(* IEC 61131-3 sources: volt/packages/volt-lsp-iec/test-corpus/lenze-mid/Device/Plc Logic/Application/Library Manager/L_OEEA_Library, 3.26.4.21 (Lenze), 47 files *)

(* ---- AXIS_REF_SIM.dut ---- *)
TYPE AXIS_REF_SIM :
STRUCT
	XENABLE : BOOL;
	XQUICKSTOP : BOOL;
	LRSETVELOCITY : LREAL;
	LRSETPOSITION : LREAL;
	XENABLED : BOOL;
	XREADY : BOOL;
	XDRIVEQSPACTIVE : BOOL;
	XERROR : BOOL;
	XWARNING : BOOL;
	EERRORID : L_IE1A_ErrorID;
	LRACTVELOCITY : LREAL;
	LRACTPOSITION : LREAL;
	XDIRECTIONPOSITIVE : BOOL;
	XDIRECTIONNEGATIVE : BOOL;
	DWDRIVEERRORID : DWORD;
	ETRAVERSINGRANGE : WORD := 1;
	LRCYCLELENGTH : LREAL := 560.0;
	LRFEEDCONSTANT : LREAL := 560.0;
	DWGEARNUMERATOR : DWORD := 77;
	DWGEARDENOMINATOR : DWORD := 6;
	XORIENTATION : BOOL := FALSE;
	EMCTRLMODE : DUT_eMctrlMode := 1;
	WNOOFHTLPERIODS : WORD := 128;
	DWHTLCOUNTERVALUE : DWORD;
	DWPOSRESOLUTION : DWORD := 65536;
	XTPRECEIVED : BOOL;
	LRTPLASTSCAN : LREAL;
	XSDOACTIVE : BOOL := TRUE;
	RDCBUSVOLTAGE : REAL;
	RMOTORCURRENT : REAL;
	RMOTORVOLTAGE : REAL;
	RMOTORSPEED : REAL;
	RMOTORFREQUENCY : REAL;
	DWERRORCODE : DWORD;
	RHEATSINKTEMP : REAL;
	RIXTLOAD : REAL;
	RIXT2LOAD : REAL;
	DWOPERATIONTIME : DWORD;
	DWSWITCHONTIME : DWORD;
	DWOPERATIONTIMECU : DWORD;
	DWOPERATIONTIMEFAN : DWORD;
END_STRUCT
END_TYPE

(* ---- DUT_EMCTRLMODE.dut ---- *)
TYPE DUT_EMCTRLMODE :
(
	OPENLOOP := 0,
	CLOSEDLOOP := 1
);
END_TYPE

(* ---- L_IE1A_ERRORID.dut ---- *)
TYPE L_IE1A_ERRORID :
(
	NOERROR := 0,
	MODULOAXISISREQUIRED := 17000,
	STARTPOSOUTOFCYCLELENGTH := 17003,
	CYCLELENGTHSHAVETOBEEQUAL := 17004,
	INVALIDDIRECTION := 17005,
	MARKSTACKLIMITREACHED := 17006,
	MAXMISSEDMARKS := 17007,
	INVALIDFOLLOWLINEACCVEL := 17008,
	INVALIDJOGGINGACCVEL := 17009,
	INVALIDSTOPDEC := 17010,
	INVALIDDIAMETER := 17011,
	TORQUEFOLLOWERNOTREADYFORMOTION := 17012,
	SPEEDFOLLOWERNOTREADYFORMOTION := 17013,
	INVALIDINVERTER := 17014,
	SDO_ACCESSFAILEDTOMOTORPARAMETERS := 17015,
	MISSEDMAPPINGPARAMETERLOWERSPEEDLIMIT := 17016,
	MISSEDMAPPINGPARAMETERUPPERSPEEDLIMIT := 17017,
	MISSEDMAPPINGPARAMETERTORQUEOFFSET := 17018,
	DANCERPOSOUTOFRANGE := 17019,
	INVALIDLIMITDANCERPOS := 17020,
	INVALIDCLUTCHPARAMETERS := 17021,
	WASNOTCALLEDDURINGMOTION := 17022,
	INVALIDNUMBEROFCAMPOINTS := 17030,
	INVALIDPATHPAR := 17032,
	INVALIDBLENDINGRADIUS := 17033,
	PATHNOTSUPPORTED := 17034,
	X_PATHLIMITPOSITIVEEXCEEDED := 17035,
	X_PATHLIMITNEGATIVEEXCEEDED := 17036,
	Y_PATHLIMITPOSITIVEEXCEEDED := 17037,
	Y_PATHLIMITNEGATIVEEXCEEDED := 17038,
	Z_PATHLIMITPOSITIVEEXCEEDED := 17039,
	Z_PATHLIMITNEGATIVEEXCEEDED := 17040,
	C_PATHLIMITPOSITIVEEXCEEDED := 17041,
	C_PATHLIMITNEGATIVEEXCEEDED := 17042,
	INVALIDPATHDATA := 17043,
	INVALIDTARGETPLC := 17047,
	MASTERISMOVING := 17100,
	INVALIDPODUCTLENGTH := 17101,
	TPSENSORNOTTEACHED := 17102,
	SLAVERECEIVEDGAPS := 17103,
	MASTERRECEIVEDGAPS := 17104,
	INTERNALERROR := 17105,
	INVALIDPARAMETERCUTTINGANGLE := 17106,
	INVALIDCUTTINGPARAMETERS := 17107,
	INVALIDCUTTINGLENGTH := 17108,
	SLAVENOTINPARKPOS := 17109,
	MASTERISREVERSING := 17110,
	INTINVALIDSELECTCAM := 17111,
	SELECTEDAXISISNOTSUPPORTED := 17112,
	AXISISNOTSUPPORTED := 17113,
	INVALIDPROFILE := 17114,
	AXISENABLEDISREQUIRED := 17115,
	CORRLIMITOUTOFCYCLELENGTH := 17116,
	CORRECTIONGREATERCORRWINDOW := 17117,
	INVALIDCNCPROGRAM := 17118,
	INVALIDGCODELINE := 17121,
	COORDSYSTEMACSNOTSUPPORTED := 17122,
	DANCERLIMITSNOTTEACHED := 17123,
	NOTREADYFORADDPROFILE := 17124,
	SLAVEPOSUPPERLIMIT := 17125,
	SLAVEPOSLOWERLIMIT := 17126,
	TARGETPOSUPPERLIMIT := 17127,
	INVALIDMARKPOSITION := 17128,
	INVALIDPOSITIONINGMODE := 17129,
	TEMPSENSORFAILURE := 17130,
	MAXCRITICALTEMPREACHED := 17131,
	INVALIDTEMPCONTROLPARAM := 17132,
	IDENTIFICATIONFAILED := 17133,
	PWMTASKCYCLEMISMATCH := 17134,
	CONCURRENTREQUESTTEMPCONTROL := 17135,
	TMNOTCALLEDINCYCLICTASK := 17136,
	TMDATABUSDISCONNECTED := 17137,
	INVALIDTMDATABUS := 17138,
	TMDATABUSCONFIGCHANGED := 17139,
	TMNOTCALLEDINMOTIONTASK := 17140,
	SLAVETMSTATESERVICE := 17141,
	COLLISIONDETECTIONDISABLED := 17142,
	COLLISIONDETECTED := 17143,
	INVALIDTMDATABUSORDER := 17144,
	CHANGEOFCONVEYORAXESNOTALLOWED := 17145,
	INVALIDSETTARGET := 17146,
	LOWERLIMITEXCEEDSUPPERLIMIT := 17147,
	SETTARGETSTACKLIMITREACHED := 17148,
	WORKPIECESTACKLIMITREACHED := 17149,
	INVALIDTRAVERSINGPROFILEPARAMETER := 17150,
	INVALIDTRAVERSINGCOILPARAMETER := 17151,
	TRAVERSINGANGULARSHIFTLIMITREACHED := 17152,
	AXESGROUPALREADYINUSE := 17153,
	UNDERVOLTAGEDCLINK := 17154,
	COUPLINGMODEREQUIRESMODULOAXIS := 17155,
	DUPLICATEDTM_ADDRESS := 17156,
	XAXISTMERROR := 17157,
	YAXISTMERROR := 17158,
	APAXISTMERROR := 17159,
	SLAVEXAXISTMERROR := 17160,
	SLAVEYAXISTMERROR := 17161,
	INVALIDMOVEPPACTIVE := 17162,
	INVALIDCONVEYORBELTPAR := 17163,
	IDENTIFICATIONDIAMETERFAILED := 17164,
	ACTDANCERPOSGTMAXDANCERPOS := 17165,
	INVALIDIDENTMAXDANCERPOS := 17166,
	INVALIDDANCERMATERIALLENGTH := 17167,
	LOADDIAMETERNOTALLOWED := 17168,
	INVALIDMASTERAXISREF := 17169,
	SYNCMODEVELACCREQUIRED := 17170,
	TEMPMAXCRITICALEXCEEDED := 17171,
	INVALIDTEMPCTRLPARAM := 17172,
	INVALIDSYNCSLAVEDIRECTION := 17173,
	MARKCORRECTIONINNEXTCYCLE := 17174,
	BASEVELOCITYNOTSUPPORTED := 17175,
	MOVEMENTBLOCKEDBYTRAINAHEAD := 17176,
	MARKDISTANCEGTZEROREQUIRED := 17177,
	INVALIDVIRTMASTERSETVELZERO := 17178,
	CONCURRENTMOTIONCMDDURINGHOMING := 17180,
	MISSINGMM_ADDRESS := 17901,
	TOOMANYMODULES := 17902,
	DUPLICATEDROOTMODULE := 17903,
	SLAVENOTFOUND := 17904,
	MISSINGAPPLICATIONREFERENCE := 17905,
	MISSINGMODULEREFERENCE := 17906,
	ERRORLISTOVERFLOW := 17907,
	ACDOWNSTRUCTINVALID := 17908,
	ACDSLAVESTRUCTINVALID := 17909,
	ACDSIZEOVERFLOW := 17910,
	COMPIDOUTOFRANGE := 17911,
	TOOMANYLEVELS := 17912,
	MMDSTRUCTINVALID := 17913,
	MODENUMBEROUTSIDERANGE := 18001,
	MODENUMBERNOTUSEDINCONFIG := 18002,
	MODECHANGENOTALLOWEDINCURRENTMODE := 18003,
	MODECHANGENOTALLOWEDINNEXTMODE := 18004,
	LI_MODENUMBEROUTSIDERANGE := 18005,
	LI_MODENUMBERNOTUSEDINCONFIG := 18006,
	LI_MODECHANGENOTALLOWEDREMOTE := 18007,
	LI_MODECHANGENOTALLOWEDINCURRENTMODE := 18008,
	LI_MODECHANGENOTALLOWEDINNEXTMODE := 18009,
	MORETHANONECOMMANDACTIVE := 18010,
	CONCURRENTCOMMAND := 18011,
	COMMANDNOTALLOWEDINCURRENTSTATE := 18012,
	LI_COMMANDSONLYINMODEPRODUCTION := 18013,
	LI_COMMANDNOTALLOWEDINREMOTE := 18014,
	LI_COMMANDNOTALLOWEDINCURRENTSTATE := 18015,
	DELAYTIMEINVALID_PT1FILTER := 19000,
	MODEINVALID_CURVE := 19002,
	MODEINVALID_COMPARE := 19003,
	MODEINVALID_CONVAXISV := 19005,
	DELAYTIMEINVALID_PROCESSCONTROLLER := 19006,
	RATETIMEINVALID_PROCESSCONTROLLER := 19007,
	RESETTIMEINVALID_PROCESSCONTROLLER := 19008,
	MODEINVALID_DELAY := 19024,
	ABORTEDBYSTARTIDENT_FRICTCOMP := 19030,
	ABORTEDBYFOLLOWERDISABLED_FRICTCOMP := 19031,
	MAXSPEEDNOTREACHED_FRICTCOMP := 19032,
	ACCTOOBIG_FRICTCOMP := 19033,
	DMINBIGGERDMAX_CALCDIAMETER := 19034,
	MAXSPEEDORMAXTORQUE_IDENTMINERTIA := 19048,
	ABORTEDBYSTARTIDENT_IDENTMINERTIA := 19049,
	ABORTEDBYFOLLOWERDISABLED_IDENTMINERTIA := 19050,
	ABORTEDBYFOLLOWERENABLED_IDENTMINERTIA := 19051,
	NMAXNOTREACHED_IDENTMINERTIA := 19052,
	MNOTREACHED_IDENTMINERTIA := 19053,
	MAXNROFTPEXCEEDED_MARKREGISTER := 19503,
	IDENTMODENOTSUPPORTED := 19801,
	MOTORRATEDSPEEDZERO := 19803,
	INERTIAMOTORZERO := 19804,
	STARTMODEINVALID := 19806,
	INVALIDEIGENFREQUENCY := 19807,
	INVALIDAMPLITUDERATIO := 19808,
	INVALIDOSCCOMPMODE := 19809,
	CHANGEOFOSCCOMPMODELOCKED := 19810,
	SDO_OTHERERROR := 20001,
	SDO_INVALIDINDEX := 20002,
	SDO_INVALIDOFFSET := 20003,
	SDO_INVALIDSIZE := 20004,
	SDO_INVALIDDATA := 20005,
	SDO_NOTREADY := 20006,
	SDO_BUSY := 20007,
	SDO_NOMEMORY := 20008,
	SDO_INVALIDPARM := 20009,
	SDO_INVALIDSTATE := 20010,
	SDO_TIMEOUT := 20011,
	SDO_INVALID_SLAVE_STATE := 20012,
	SDO_LINK_DISCONNECTED := 20013,
	SDO_ALL_CANNELS_BUSY := 20015,
	SDO_ABORTCODE_TOGGLE := 20020,
	SDO_ABORTCODE_TIMEOUT := 20021,
	SDO_ABORTCODE_CCS_SCS := 20022,
	SDO_ABORTCODE_BLK_SIZE := 20023,
	SDO_ABORTCODE_SEQNO := 20024,
	SDO_ABORTCODE_CRC := 20025,
	SDO_ABORTCODE_MEMORY := 20026,
	SDO_ABORTCODE_ACCESS := 20027,
	SDO_ABORTCODE_WRITEONLY := 20028,
	SDO_ABORTCODE_READONLY := 20029,
	SDO_ABORTCODE_INDEX := 20030,
	SDO_ABORTCODE_PDO_MAP := 20031,
	SDO_ABORTCODE_PDO_LEN := 20032,
	SDO_ABORTCODE_P_INCOMP := 20033,
	SDO_ABORTCODE_I_INCOMP := 20034,
	SDO_ABORTCODE_HARDWARE := 20035,
	SDO_ABORTCODE_DATA_SIZE := 20036,
	SDO_ABORTCODE_DATA_SIZE1 := 20037,
	SDO_ABORTCODE_DATA_SIZE2 := 20038,
	SDO_ABORTCODE_OFFSET := 20039,
	SDO_ABORTCODE_DATA_RANGE := 20040,
	SDO_ABORTCODE_DATA_RANGE1 := 20041,
	SDO_ABORTCODE_DATA_RANGE2 := 20042,
	SDO_ABORTCODE_MINMAX := 20043,
	SDO_ABORTCODE_GENERAL := 20044,
	SDO_ABORTCODE_TRANSFER := 20045,
	SDO_ABORTCODE_TRANSFER1 := 20046,
	SDO_ABORTCODE_TRANSFER2 := 20047,
	SDO_ABORTCODE_DICTIONARY := 20048,
	SDO_ABORTCODE_UNKNOWN := 20049,
	NOAXISREF := 20301,
	NOPARAMETER := 20302,
	NOVALIDPARAM := 20303,
	NOVALIDAXISSTATE := 20304,
	NOBOOLPARAM := 20305,
	SWLIMITPOS := 20306,
	SWLIMITNEG := 20307,
	NOVALID_MC_SOURCE := 20308,
	NOSETVALUESAVAILABLE := 20309,
	POWERFAILDURINGOPERATION := 20310,
	NOTREADYFORMOTION := 20311,
	POSSWLIMITREACHED := 20312,
	NEGSWLIMITREACHED := 20313,
	NOVALIDTPSOURCE := 20314,
	NOVALIDTPNUMBER := 20315,
	TPALREADYACTIVE := 20316,
	NOTTPSUPPORTED := 20317,
	NOTPACTIVE := 20318,
	NOEXTPINPUT := 20319,
	NOVALIDACCELERATION := 20320,
	NOVALIDDECELERATION := 20321,
	NOVALIDVELOCITY := 20322,
	ARITHMETICERROR := 20323,
	NOTAPPLICABLE := 20324,
	VELOCITYLIMITED := 20325,
	ACCELERATIONLIMITED := 20326,
	JERKLIMITED := 20327,
	TARGETOUTSIDESWLIMIT := 20328,
	NOVALIDACCELERATION_MOVEABSOLUTE := 20330,
	NOVALIDDECELERATION_MOVEABSOLUTE := 20331,
	NOVALIDVELOCITY_MOVEABSOLUTE := 20332,
	ARITHMETICERROR_MOVEABSOLUTE := 20333,
	NOTAPPLICABLE_MOVEABSOLUTE := 20334,
	VELOCITYLIMITED_MOVEABSOLUTE := 20335,
	ACCELERATIONLIMITED_MOVEABSOLUTE := 20336,
	JERKLIMITED_MOVEABSOLUTE := 20337,
	TARGETOUTSIDESWLIMIT_MOVEABSOLUTE := 20338,
	NOVALIDACCELERATION_MOVEADDITIVE := 20340,
	NOVALIDDECELERATION_MOVEADDITIVE := 20341,
	NOVALIDVELOCITY_MOVEADDITIVE := 20342,
	ARITHMETICERROR_MOVEADDITIVE := 20343,
	NOTAPPLICABLE_MOVEADDITIVE := 20344,
	VELOCITYLIMITED_MOVEADDITIVE := 20345,
	ACCELERATIONLIMITED_MOVEADDITIVE := 20346,
	JERKLIMITED_MOVEADDITIVE := 20347,
	TARGETOUTSIDESWLIMIT_MOVEADDITIVE := 20348,
	NOVALIDACCELERATION_MOVECONTAB := 20350,
	NOVALIDDECELERATION_MOVECONTAB := 20351,
	NOVALIDVELOCITY_MOVECONTAB := 20352,
	ARITHMETICERROR_MOVECONTAB := 20353,
	NOTAPPLICABLE_MOVECONTAB := 20354,
	VELOCITYLIMITED_MOVECONTAB := 20355,
	ACCELERATIONLIMITED_MOVECONTAB := 20356,
	JERKLIMITED_MOVECONTAB := 20357,
	TARGETOUTSIDESWLIMIT_MOVECONTAB := 20358,
	NOVALIDACCELERATION_MOVECONTREL := 20360,
	NOVALIDDECELERATION_MOVECONTREL := 20361,
	NOVALIDVELOCITY_MOVECONTREL := 20362,
	ARITHMETICERROR_MOVECONTREL := 20363,
	NOTAPPLICABLE_MOVECONTREL := 20364,
	VELOCITYLIMITED_MOVECONTREL := 20365,
	ACCELERATIONLIMITED_MOVECONTREL := 20366,
	JERKLIMITED_MOVECONTREL := 20367,
	TARGETOUTSIDESWLIMIT_MOVECONTREL := 20368,
	NOVALIDACCELERATION_MOVERELATIVE := 20370,
	NOVALIDDECELERATION_MOVERELATIVE := 20371,
	NOVALIDVELOCITY_MOVERELATIVE := 20372,
	ARITHMETICERROR_MOVERELATIVE := 20373,
	NOTAPPLICABLE_MOVERELATIVE := 20374,
	VELOCITYLIMITED_MOVERELATIVE := 20375,
	ACCELERATIONLIMITED_MOVERELATIVE := 20376,
	JERKLIMITED_MOVERELATIVE := 20377,
	TARGETOUTSIDESWLIMIT_MOVERELATIVE := 20378,
	NOVALIDACCELERATION_MOVESUPERIMP := 20380,
	NOVALIDDECELERATION_MOVESUPERIMP := 20381,
	NOVALIDVELOCITY_MOVESUPERIMP := 20382,
	ARITHMETICERROR_MOVESUPERIMP := 20383,
	NOTAPPLICABLE_MOVESUPERIMP := 20384,
	VELOCITYLIMITED_MOVESUPERIMP := 20385,
	ACCELERATIONLIMITED_MOVESUPERIMP := 20386,
	JERKLIMITED_MOVESUPERIMP := 20387,
	TARGETOUTSIDESWLIMIT_MOVESUPERIMP := 20388,
	NOVALIDACCELERATION_MOVEVELOCITY := 20390,
	NOVALIDDECELERATION_MOVEVELOCITY := 20391,
	NOVALIDVELOCITY_MOVEVELOCITY := 20392,
	ARITHMETICERROR_MOVEVELOCITY := 20393,
	NOTAPPLICABLE_MOVEVELOCITY := 20394,
	VELOCITYLIMITED_MOVEVELOCITY := 20395,
	ACCELERATIONLIMITED_MOVEVELOCITY := 20396,
	JERKLIMITED_MOVEVELOCITY := 20397,
	TARGETOUTSIDESWLIMIT_MOVEVELOCITY := 20398,
	NOVALIDDECELERATION_HALT := 20401,
	ARITHMETICERROR_HALT := 20403,
	ACCELERATIONLIMITED_HALT := 20406,
	JERKLIMITED_HALT := 20407,
	NOVALIDDECELERATION_STOP := 20411,
	ARITHMETICERROR_STOP := 20413,
	ACCELERATIONLIMITED_STOP := 20416,
	JERKLIMITED_STOP := 20417,
	NOVALIDDIRECTION := 20430,
	NOVALIDBUFFERMODE := 20431,
	DIRECTIONDISABLED := 20432,
	BLOCKEDBYAXISSTATE := 20433,
	NOVALIDOVERRIDE := 20434,
	CONCURRENT_MC_POWER := 20435,
	CONCURRENT_SETQUICKSTOP := 20436,
	DRIVE_PDO_INTERFACE_DISABLED := 20499,
	HWLIMITPOS := 20500,
	HWLIMITNEG := 20501,
	FOLLOWINGERROR1 := 20502,
	FOLLOWINGERROR2 := 20503,
	COMMUNICATIONFAIL := 20504,
	AXISINITFAIL := 20505,
	COMMTIMOUT := 20506,
	MASTERRESTARTFAIL := 20507,
	NOTREADYFORREINIT := 20508,
	ERRORDURINGINIT := 20509,
	SWITCHONNOTPOSSIBLE := 20510,
	DRIVEERROR := 20511,
	HOME_NOAUXPARAMETERS := 20512,
	HOME_MODENOTSUPPORTEDBYAXIS := 20513,
	HOME_MODEUNKNOWN := 20514,
	HOME_NOAUXTRIGGERINPUT := 20515,
	HOME_UNKNOWNTPCONFIG := 20516,
	HOME_WRITEHOMEPARAMETER := 20518,
	HOME_ERRORWHILEHOMING := 20519,
	HOME_ARITHMETICERROR := 20520,
	HOME_TORQUELIMNOTMAPPED := 20521,
	HOME_INVALIDVELACC := 20522,
	HOMETPEDGESETTINGNOTSUPPORTED := 20523,
	RESETDRIVEERRORFAILED := 20525,
	APPLICATIONERROR := 20526,
	APPLICATIONWARNING := 20527,
	BRAKE_POSITIONDRIFT := 20529,
	BRAKE_INVALIDMODE := 20530,
	BRAKE_TIMEOUTPRECONTROL := 20531,
	BRAKE_INVALIDBRAKESTATE := 20532,
	FAST_IO_OUT_WRONGOUTPUTSEL := 20533,
	FAST_IO_OUT_NOFREEENCODERAXIS := 20534,
	FAST_IO_OUT_FREEENCODERAXISWRONGPARAMETER := 20535,
	FAST_IO_OUT_MAPPINGFAULT := 20536,
	FAST_IO_OUT_FIFOOVERFLOW := 20537,
	TP_SELECT := 20538,
	TP_MODE := 20539,
	TP_EDGENOTAVAILABLE := 20541,
	TP_CHANNELNOTFREE := 20542,
	TP_MAPPINGFAULT := 20543,
	TP_INTERNALCHANNELNOTFREE := 20544,
	TP_TIMEOUT := 20545,
	TP_COMMUNICATIONERROR := 20546,
	TP_SIGNAL := 20547,
	TP_NOFREEENCODERAXIS := 20548,
	TP_PARAMETERRISINGEDGEWRONGVALUE := 20550,
	TP_PARAMETERFALLINGRISINGEDGEWRONGVALUE := 20551,
	TP_INTERNALERROR := 20552,
	SETVALUESGTMAXAPPVALUES := 20600,
	SETVALUESINCONSISTENT := 20601,
	POSDIFFGTHALFCYCLELENGTH := 20602,
	INVALIDTASKCYCLETIME := 20603,
	INIT_WRITEERRORSDO := 20650,
	INIT_READERRORSDO := 20651,
	INIT_MAXTASKTIME := 20652,
	INIT_TORQUEREFISZERO := 20653,
	INIT_MOTORRATEDSPEEDISZERO := 20654,
	INIT_REVISIONNOTVALID := 20655,
	INIT_ENCCOUNTNOTVALID := 20656,
	INIT_ENCREVNOTVALID := 20657,
	INIT_ENCCRCNOTVALID := 20658,
	INIT_ENCABSPOSNOTAVAILABLE := 20659,
	CONTROLLERFIRMWARENOTCOMPATIBLE := 20660,
	INVALIDMODE := 20661,
	ENCBPB_INIT_FAILED := 20662,
	LEDNOTSUPPORTEDBYDEVICE := 20663,
	INVALIDGEARFACTOR := 20664,
	POSOUTOFCYCLELENGTH := 20665,
	CYCLELENGTHINVALID_ADDOFFSETCYCLIC := 20666,
	POSININVALID_ADDOFFSETCYCLIC := 20667,
	CYCLELENGTHINVALID_ZERODETECT := 20668,
	POSININVALID_ZERODETECT := 20669,
	STARTPOSINVALID_INTEGRATEAXIS := 20670,
	INVALIDINPUTJOGPOSJOGNEG := 20671,
	VALUEOUTOFRANGE := 20672,
	STATENOTEQUALDISABLED := 20673,
	INVALIDINPUT_BRAKETEST := 20674,
	ALREADYACTIVE_BRAKETEST := 20675,
	INVALIDINPUT_BRAKEGRINDIN := 20676,
	ALREADYACTIVE_GRINDIN := 20677,
	INVALIDCONTROLMODE := 20678,
	VIRTUALAXISNOTSUPPORTED := 20679,
	AXISNOTDISABLED := 20680,
	INVALIDFEEDCONSTANT := 20681,
	INVALIDTRAVERSINGRANGE := 20682,
	INVALIDCYCLELENGTH := 20683,
	INVALIDPOSRESOLUTION := 20684,
	TORQUELIMTOOLARGE := 20685,
	TORQUELIMLESSTHANZERO := 20686,
	ENCSIGNALINVALID := 20687,
	ENCSIGNALGTMEASURINGRANGE := 20688,
	INVALIDENCMEASURINGRANGE := 20689,
	DRIVESTOACTIVE := 20690,
	DRIVECINHACTIVE := 20691,
	INVALIDSWLIMITS := 20692,
	NOVALIDJERK := 20693,
	MISSEDMAPPINGPARAMETERVLTARGETVEL := 20694,
	MISSEDMAPPINGPARAMETERVLACTUALVEL := 20695,
	AXISNOTHOMED := 20696,
	AXISNOTINSIMPLEMODE := 20697,
	AXISINSIMPLEMODE := 20698,
	FUNCTIONNOTSUPPORTEDBYAXIS := 20699,
	EXECUTIONINDEXALREADYINUSE := 20700,
	SS1ACTIVE := 20701,
	SS2ACTIVE := 20702,
	VELOCITYLIMITEDBYSLS1 := 20703,
	VELOCITYLIMITEDBYSLS2 := 20704,
	VELOCITYLIMITEDBYSLS3 := 20705,
	VELOCITYLIMITEDBYSLS4 := 20706,
	INVALIDEXECUTIONINDEX := 20707,
	INVALIDFILTERDEPTH := 20708,
	PARAMSETFAILEDJOGVEL := 20709,
	PARAMSETFAILEDJOGACC := 20710,
	PARAMSETFAILEDJOGDEC := 20711,
	PARAMSETFAILEDJOGJERK := 20712,
	PARAMSETFAILEDHALTDEC := 20713,
	PARAMSETFAILEDHALTJERK := 20714,
	PARAMSETFAILEDQSPAPPLDEC := 20715,
	PARAMSETFAILEDQSPAPPLJERK := 20716,
	PARAMSETFAILEDHOMEPOSITION := 20717,
	PARAMSETFAILEDHOMEMODE := 20718,
	PARAMSETFAILEDHOMESTOPMODE := 20719,
	PARAMSETFAILEDHOMETARGETPOSITION := 20720,
	PARAMSETFAILEDHOMEVELOCITY1 := 20721,
	PARAMSETFAILEDHOMEVELOCITY2 := 20722,
	PARAMSETFAILEDHOMEACCELERATION1 := 20723,
	PARAMSETFAILEDHOMEACCELERATION2 := 20724,
	PARAMSETFAILEDHOMEJERK := 20725,
	PARAMSETFAILEDHOMETORQUELIMIT := 20726,
	PARAMSETFAILEDHOMETORQUETIME := 20727,
	PARAMSETFAILEDHOMETPCONFIG := 20728,
	PARAMSETFAILEDDRIVEHOMEMODE := 20729,
	PARAMREADFAILED := 20730,
	PARAMROLLBACKFAILED := 20731,
	POSCTRLNOTSUPPORTED := 20732,
	TORQUECTRLNOTSUPPORTED := 20733,
	SETPOSITIONINPDOREQUIRED := 20734,
	SETVELOCITYINPDOREQUIRED := 20735,
	SETTORQUEINPDOREQUIRED := 20736,
	UPPERSPEEDLIMINPDOREQUIRED := 20737,
	LOWERSPEEDLIMINPDOREQUIRED := 20738,
	ACTPOSITIONINPDOREQUIRED := 20739,
	BRAKEGRINDININVALIDPOSITIONLIMITS := 20740,
	BRAKEGRINDINSTARTPOSOUTSIDEPOSLIM := 20741,
	BRAKEGRINDINDISTANCENOTSUFFICIENT := 20742,
	SAFETYNOTSUPPORTEDBYDRIVE := 20743,
	SAFETYCONTROLWORDINPDOREQUIRED := 20744,
	SETPOSITIONONSLAVEAXISNOTALLOWED := 20745,
	ENCODERVELOCITYGTMAXVELOCITY := 20746,
	INVALIDENCODERSIGNAL := 20747,
	DRIVESAFEBRAKECTRLACTIVE := 20748,
	POSRECONSTRDATAINKONSISTENT := 20750,
	POSRECONSTRHOMEPOSAVAILABLENOTACTIVE := 20751,
	POSRECONSTRNOTACTIVATED := 20752,
	POSRECONSTRAXISWASVIRTUAL := 20753,
	POSRECONSTRORIENTATIONCHANGED := 20754,
	POSRECONSTRTRAVERSINGRANGECHANGED := 20755,
	POSRECONSTRCYCLELENGTHCHANGED := 20756,
	POSRECONSTRUNITFACTORCHANGED := 20757,
	POSRECONSTRRESETBYENCERROR := 20758,
	POSRECONSTRRESETBYFDBCHANGED := 20759,
	POSRECONSTRENCCRCCHANGED := 20760,
	POSRECONSTRNOFDBPOSAVAILABLE := 20761,
	POSRECONSTRABSENCREQUIRED := 20762,
	POSRECONSTRDATAVERSIONCHANGED := 20763,
	POSRECONSTRNODATAAVAILABLE := 20764,
	POSRECONSTRNOMEMORYAVAILABLE := 20765,
	POSRECONSTRPOSOUTSIDERESTORETRESHOLD := 20766,
	POSRECONSTRRESETBYFDBOPENCIRC := 20767,
	MAINAXISNOTREADY := 21001,
	GROUPSTATEUNDEFINED := 21002,
	AXISDISABLED := 21003,
	TRANSFORMATIONERROR := 21004,
	AXISINERRORSTOP := 21005,
	AXISLIMITVIOLATIONMAINAXIS := 21006,
	AXISLIMITVIOLATIONREALAXIS := 21007,
	AXISLIMITVIOLATIONPASSIVEAXIS := 21008,
	REALAXISDISABLED := 21009,
	NOVALIDPATHCOICE_MOVECIRCABS := 21010,
	NOVALIDCIRCMODE_MOVECIRCABS := 21011,
	NOVALIDTRANSITIONPARAMETER_MOVECIRCABS := 21012,
	NOVALIDVELOCITY_MOVECIRCABS := 21013,
	NOVALIDACCELERATION_MOVECIRCABS := 21014,
	NOVALIDDECELERATION_MOVECIRCABS := 21015,
	NOVALIDJERK_MOVECIRCABS := 21016,
	TARGETOUTSIDESWLIMITSPASSIVEJOINTS_MOVECIRCABS := 21017,
	TARGETOUTSIDESWLIMITSMAINAXISX_MOVECIRCABS := 21018,
	TARGETOUTSIDESWLIMITSMAINAXISY_MOVECIRCABS := 21019,
	TARGETOUTSIDESWLIMITSMAINAXISZ_MOVECIRCABS := 21020,
	TARGETOUTSIDESWLIMITSMAINAXISA_MOVECIRCABS := 21021,
	TARGETOUTSIDESWLIMITSMAINAXISB_MOVECIRCABS := 21022,
	TARGETOUTSIDESWLIMITSMAINAXISC_MOVECIRCABS := 21023,
	TARGETOUTSIDESWLIMITSREALAXIS1_MOVECIRCABS := 21024,
	TARGETOUTSIDESWLIMITSREALAXIS2_MOVECIRCABS := 21025,
	TARGETOUTSIDESWLIMITSREALAXIS3_MOVECIRCABS := 21026,
	TARGETOUTSIDESWLIMITSREALAXIS4_MOVECIRCABS := 21027,
	TARGETOUTSIDESWLIMITSREALAXIS5_MOVECIRCABS := 21028,
	TARGETOUTSIDESWLIMITSREALAXIS6_MOVECIRCABS := 21029,
	TARGETOUTSIDESWLIMITSAUXAXIS1_MOVECIRCABS := 21030,
	TARGETOUTSIDESWLIMITSAUXAXIS2_MOVECIRCABS := 21031,
	TARGETOUTSIDESWLIMITSAUXAXIS3_MOVECIRCABS := 21032,
	TARGETOUTSIDESWLIMITSAUXAXIS4_MOVECIRCABS := 21033,
	TARGETOUTSIDESWLIMITSAUXAXIS5_MOVECIRCABS := 21034,
	TARGETOUTSIDESWLIMITSAUXAXIS6_MOVECIRCABS := 21035,
	TARGETTRANSFORMATIONERROR_MOVECIRCABS := 21036,
	TARGETSINGULARPOS_MOVECIRCABS := 21037,
	BORDEROUTSIDESWLIMITSPASSIVEJOINTS_MOVECIRCABS := 21038,
	BORDEROUTSIDESWLIMITSMAINAXISX_MOVECIRCABS := 21039,
	BORDEROUTSIDESWLIMITSMAINAXISY_MOVECIRCABS := 21040,
	BORDEROUTSIDESWLIMITSMAINAXISZ_MOVECIRCABS := 21041,
	BORDEROUTSIDESWLIMITSMAINAXISA_MOVECIRCABS := 21042,
	BORDEROUTSIDESWLIMITSMAINAXISB_MOVECIRCABS := 21043,
	BORDEROUTSIDESWLIMITSMAINAXISC_MOVECIRCABS := 21044,
	BORDEROUTSIDESWLIMITSREALAXIS1_MOVECIRCABS := 21045,
	BORDEROUTSIDESWLIMITSREALAXIS2_MOVECIRCABS := 21046,
	BORDEROUTSIDESWLIMITSREALAXIS3_MOVECIRCABS := 21047,
	BORDEROUTSIDESWLIMITSREALAXIS4_MOVECIRCABS := 21048,
	BORDEROUTSIDESWLIMITSREALAXIS5_MOVECIRCABS := 21049,
	BORDEROUTSIDESWLIMITSREALAXIS6_MOVECIRCABS := 21050,
	BORDEROUTSIDESWLIMITSAUXAXIS1_MOVECIRCABS := 21051,
	BORDEROUTSIDESWLIMITSAUXAXIS2_MOVECIRCABS := 21052,
	BORDEROUTSIDESWLIMITSAUXAXIS3_MOVECIRCABS := 21053,
	BORDEROUTSIDESWLIMITSAUXAXIS4_MOVECIRCABS := 21054,
	BORDEROUTSIDESWLIMITSAUXAXIS5_MOVECIRCABS := 21055,
	BORDEROUTSIDESWLIMITSAUXAXIS6_MOVECIRCABS := 21056,
	BORDERTRANSFORMATIONERROR_MOVECIRCABS := 21057,
	BORDERSINGULARPOS_MOVECIRCABS := 21058,
	ILLEGALPARAMETER_MOVECIRCABS := 21059,
	NOVALIDPATHCOICE_MOVECIRCREL := 21060,
	NOVALIDCIRCMODE_MOVECIRCREL := 21061,
	NOVALIDTRANSITIONPARAMETER_MOVECIRCREL := 21062,
	NOVALIDVELOCITY_MOVECIRCREL := 21063,
	NOVALIDACCELERATION_MOVECIRCREL := 21064,
	NOVALIDDECELERATION_MOVECIRCREL := 21065,
	NOVALIDJERK_MOVECIRCREL := 21066,
	TARGETOUTSIDESWLIMITSPASSIVEJOINTS_MOVECIRCREL := 21067,
	TARGETOUTSIDESWLIMITSMAINAXISX_MOVECIRCREL := 21068,
	TARGETOUTSIDESWLIMITSMAINAXISY_MOVECIRCREL := 21069,
	TARGETOUTSIDESWLIMITSMAINAXISZ_MOVECIRCREL := 21070,
	TARGETOUTSIDESWLIMITSMAINAXISA_MOVECIRCREL := 21071,
	TARGETOUTSIDESWLIMITSMAINAXISB_MOVECIRCREL := 21072,
	TARGETOUTSIDESWLIMITSMAINAXISC_MOVECIRCREL := 21073,
	TARGETOUTSIDESWLIMITSREALAXIS1_MOVECIRCREL := 21074,
	TARGETOUTSIDESWLIMITSREALAXIS2_MOVECIRCREL := 21075,
	TARGETOUTSIDESWLIMITSREALAXIS3_MOVECIRCREL := 21076,
	TARGETOUTSIDESWLIMITSREALAXIS4_MOVECIRCREL := 21077,
	TARGETOUTSIDESWLIMITSREALAXIS5_MOVECIRCREL := 21078,
	TARGETOUTSIDESWLIMITSREALAXIS6_MOVECIRCREL := 21079,
	TARGETOUTSIDESWLIMITSAUXAXIS1_MOVECIRCREL := 21080,
	TARGETOUTSIDESWLIMITSAUXAXIS2_MOVECIRCREL := 21081,
	TARGETOUTSIDESWLIMITSAUXAXIS3_MOVECIRCREL := 21082,
	TARGETOUTSIDESWLIMITSAUXAXIS4_MOVECIRCREL := 21083,
	TARGETOUTSIDESWLIMITSAUXAXIS5_MOVECIRCREL := 21084,
	TARGETOUTSIDESWLIMITSAUXAXIS6_MOVECIRCREL := 21085,
	TARGETTRANSFORMATIONERROR_MOVECIRCREL := 21086,
	TARGETSINGULARPOS_MOVECIRCREL := 21087,
	BORDEROUTSIDESWLIMITSPASSIVEJOINTS_MOVECIRCREL := 21088,
	BORDEROUTSIDESWLIMITSMAINAXISX_MOVECIRCREL := 21089,
	BORDEROUTSIDESWLIMITSMAINAXISY_MOVECIRCREL := 21090,
	BORDEROUTSIDESWLIMITSMAINAXISZ_MOVECIRCREL := 21091,
	BORDEROUTSIDESWLIMITSMAINAXISA_MOVECIRCREL := 21092,
	BORDEROUTSIDESWLIMITSMAINAXISB_MOVECIRCREL := 21093,
	BORDEROUTSIDESWLIMITSMAINAXISC_MOVECIRCREL := 21094,
	BORDEROUTSIDESWLIMITSREALAXIS1_MOVECIRCREL := 21095,
	BORDEROUTSIDESWLIMITSREALAXIS2_MOVECIRCREL := 21096,
	BORDEROUTSIDESWLIMITSREALAXIS3_MOVECIRCREL := 21097,
	BORDEROUTSIDESWLIMITSREALAXIS4_MOVECIRCREL := 21098,
	BORDEROUTSIDESWLIMITSREALAXIS5_MOVECIRCREL := 21099,
	BORDEROUTSIDESWLIMITSREALAXIS6_MOVECIRCREL := 21100,
	BORDEROUTSIDESWLIMITSAUXAXIS1_MOVECIRCREL := 21101,
	BORDEROUTSIDESWLIMITSAUXAXIS2_MOVECIRCREL := 21102,
	BORDEROUTSIDESWLIMITSAUXAXIS3_MOVECIRCREL := 21103,
	BORDEROUTSIDESWLIMITSAUXAXIS4_MOVECIRCREL := 21104,
	BORDEROUTSIDESWLIMITSAUXAXIS5_MOVECIRCREL := 21105,
	BORDEROUTSIDESWLIMITSAUXAXIS6_MOVECIRCREL := 21106,
	BORDERTRANSFORMATIONERROR_MOVECIRCREL := 21107,
	BORDERSINGULARPOS_MOVECIRCREL := 21108,
	ILLEGALPARAMETER_MOVECIRCREL := 21109,
	NOVALIDTRANSITIONPARAMETER_MOVELINABS := 21110,
	NOVALIDVELOCITY_MOVELINABS := 21111,
	NOVALIDACCELERATION_MOVELINABS := 21112,
	NOVALIDDECELERATION_MOVELINABS := 21113,
	NOVALIDJERK_MOVELINABS := 21114,
	TARGETOUTSIDESWLIMITSPASSIVEJOINTS_MOVELINABS := 21115,
	TARGETOUTSIDESWLIMITSMAINAXISX_MOVELINABS := 21116,
	TARGETOUTSIDESWLIMITSMAINAXISY_MOVELINABS := 21117,
	TARGETOUTSIDESWLIMITSMAINAXISZ_MOVELINABS := 21118,
	TARGETOUTSIDESWLIMITSMAINAXISA_MOVELINABS := 21119,
	TARGETOUTSIDESWLIMITSMAINAXISB_MOVELINABS := 21120,
	TARGETOUTSIDESWLIMITSMAINAXISC_MOVELINABS := 21121,
	TARGETOUTSIDESWLIMITSREALAXIS1_MOVELINABS := 21122,
	TARGETOUTSIDESWLIMITSREALAXIS2_MOVELINABS := 21123,
	TARGETOUTSIDESWLIMITSREALAXIS3_MOVELINABS := 21124,
	TARGETOUTSIDESWLIMITSREALAXIS4_MOVELINABS := 21125,
	TARGETOUTSIDESWLIMITSREALAXIS5_MOVELINABS := 21126,
	TARGETOUTSIDESWLIMITSREALAXIS6_MOVELINABS := 21127,
	TARGETOUTSIDESWLIMITSAUXAXIS1_MOVELINABS := 21128,
	TARGETOUTSIDESWLIMITSAUXAXIS2_MOVELINABS := 21129,
	TARGETOUTSIDESWLIMITSAUXAXIS3_MOVELINABS := 21130,
	TARGETOUTSIDESWLIMITSAUXAXIS4_MOVELINABS := 21131,
	TARGETOUTSIDESWLIMITSAUXAXIS5_MOVELINABS := 21132,
	TARGETOUTSIDESWLIMITSAUXAXIS6_MOVELINABS := 21133,
	TARGETTRANSFORMATIONERROR_MOVELINABS := 21134,
	TARGETSINGULARPOS_MOVELINABS := 21135,
	ILLEGALPARAMETER_MOVELINABS := 21136,
	NOVALIDTRANSITIONPARAMETER_MOVELINREL := 21137,
	NOVALIDVELOCITY_MOVELINREL := 21138,
	NOVALIDACCELERATION_MOVELINREL := 21139,
	NOVALIDDECELERATION_MOVELINREL := 21140,
	NOVALIDJERK_MOVELINREL := 21141,
	TARGETOUTSIDESWLIMITSPASSIVEJOINTS_MOVELINREL := 21142,
	TARGETOUTSIDESWLIMITSMAINAXISX_MOVELINREL := 21143,
	TARGETOUTSIDESWLIMITSMAINAXISY_MOVELINREL := 21144,
	TARGETOUTSIDESWLIMITSMAINAXISZ_MOVELINREL := 21145,
	TARGETOUTSIDESWLIMITSMAINAXISA_MOVELINREL := 21146,
	TARGETOUTSIDESWLIMITSMAINAXISB_MOVELINREL := 21147,
	TARGETOUTSIDESWLIMITSMAINAXISC_MOVELINREL := 21148,
	TARGETOUTSIDESWLIMITSREALAXIS1_MOVELINREL := 21149,
	TARGETOUTSIDESWLIMITSREALAXIS2_MOVELINREL := 21150,
	TARGETOUTSIDESWLIMITSREALAXIS3_MOVELINREL := 21151,
	TARGETOUTSIDESWLIMITSREALAXIS4_MOVELINREL := 21152,
	TARGETOUTSIDESWLIMITSREALAXIS5_MOVELINREL := 21153,
	TARGETOUTSIDESWLIMITSREALAXIS6_MOVELINREL := 21154,
	TARGETOUTSIDESWLIMITSAUXAXIS1_MOVELINREL := 21155,
	TARGETOUTSIDESWLIMITSAUXAXIS2_MOVELINREL := 21156,
	TARGETOUTSIDESWLIMITSAUXAXIS3_MOVELINREL := 21157,
	TARGETOUTSIDESWLIMITSAUXAXIS4_MOVELINREL := 21158,
	TARGETOUTSIDESWLIMITSAUXAXIS5_MOVELINREL := 21159,
	TARGETOUTSIDESWLIMITSAUXAXIS6_MOVELINREL := 21160,
	TARGETTRANSFORMATIONERROR_MOVELINREL := 21161,
	TARGETSINGULARPOS_MOVELINREL := 21162,
	ILLEGALPARAMETER_MOVELINREL := 21163,
	NOVALIDTRANSITIONPARAMETER_MOVEDIRABS := 21164,
	NOVALIDVELOCITY_MOVEDIRABS := 21165,
	NOVALIDACCELERATION_MOVEDIRABS := 21166,
	NOVALIDDECELERATION_MOVEDIRABS := 21167,
	NOVALIDJERK_MOVEDIRABS := 21168,
	TARGETOUTSIDESWLIMITSPASSIVEJOINTS_MOVEDIRABS := 21169,
	TARGETOUTSIDESWLIMITSMAINAXISX_MOVEDIRABS := 21170,
	TARGETOUTSIDESWLIMITSMAINAXISY_MOVEDIRABS := 21171,
	TARGETOUTSIDESWLIMITSMAINAXISZ_MOVEDIRABS := 21172,
	TARGETOUTSIDESWLIMITSMAINAXISA_MOVEDIRABS := 21173,
	TARGETOUTSIDESWLIMITSMAINAXISB_MOVEDIRABS := 21174,
	TARGETOUTSIDESWLIMITSMAINAXISC_MOVEDIRABS := 21175,
	TARGETOUTSIDESWLIMITSREALAXIS1_MOVEDIRABS := 21176,
	TARGETOUTSIDESWLIMITSREALAXIS2_MOVEDIRABS := 21177,
	TARGETOUTSIDESWLIMITSREALAXIS3_MOVEDIRABS := 21178,
	TARGETOUTSIDESWLIMITSREALAXIS4_MOVEDIRABS := 21179,
	TARGETOUTSIDESWLIMITSREALAXIS5_MOVEDIRABS := 21180,
	TARGETOUTSIDESWLIMITSREALAXIS6_MOVEDIRABS := 21181,
	TARGETOUTSIDESWLIMITSAUXAXIS1_MOVEDIRABS := 21182,
	TARGETOUTSIDESWLIMITSAUXAXIS2_MOVEDIRABS := 21183,
	TARGETOUTSIDESWLIMITSAUXAXIS3_MOVEDIRABS := 21184,
	TARGETOUTSIDESWLIMITSAUXAXIS4_MOVEDIRABS := 21185,
	TARGETOUTSIDESWLIMITSAUXAXIS5_MOVEDIRABS := 21186,
	TARGETOUTSIDESWLIMITSAUXAXIS6_MOVEDIRABS := 21187,
	TARGETTRANSFORMATIONERROR_MOVEDIRABS := 21188,
	ILLEGALPARAMETER_MOVEDIRABS := 21189,
	NOVALIDTRANSITIONPARAMETER_MOVEDIRREL := 21190,
	NOVALIDVELOCITY_MOVEDIRREL := 21191,
	NOVALIDACCELERATION_MOVEDIRREL := 21192,
	NOVALIDDECELERATION_MOVEDIRREL := 21193,
	NOVALIDJERK_MOVEDIRREL := 21194,
	TARGETOUTSIDESWLIMITSPASSIVEJOINTS_MOVEDIRREL := 21195,
	TARGETOUTSIDESWLIMITSMAINAXISX_MOVEDIRREL := 21196,
	TARGETOUTSIDESWLIMITSMAINAXISY_MOVEDIRREL := 21197,
	TARGETOUTSIDESWLIMITSMAINAXISZ_MOVEDIRREL := 21198,
	TARGETOUTSIDESWLIMITSMAINAXISA_MOVEDIRREL := 21199,
	TARGETOUTSIDESWLIMITSMAINAXISB_MOVEDIRREL := 21200,
	TARGETOUTSIDESWLIMITSMAINAXISC_MOVEDIRREL := 21201,
	TARGETOUTSIDESWLIMITSREALAXIS1_MOVEDIRREL := 21202,
	TARGETOUTSIDESWLIMITSREALAXIS2_MOVEDIRREL := 21203,
	TARGETOUTSIDESWLIMITSREALAXIS3_MOVEDIRREL := 21204,
	TARGETOUTSIDESWLIMITSREALAXIS4_MOVEDIRREL := 21205,
	TARGETOUTSIDESWLIMITSREALAXIS5_MOVEDIRREL := 21206,
	TARGETOUTSIDESWLIMITSREALAXIS6_MOVEDIRREL := 21207,
	TARGETOUTSIDESWLIMITSAUXAXIS1_MOVEDIRREL := 21208,
	TARGETOUTSIDESWLIMITSAUXAXIS2_MOVEDIRREL := 21209,
	TARGETOUTSIDESWLIMITSAUXAXIS3_MOVEDIRREL := 21210,
	TARGETOUTSIDESWLIMITSAUXAXIS4_MOVEDIRREL := 21211,
	TARGETOUTSIDESWLIMITSAUXAXIS5_MOVEDIRREL := 21212,
	TARGETOUTSIDESWLIMITSAUXAXIS6_MOVEDIRREL := 21213,
	TARGETTRANSFORMATIONERROR_MOVEDIRREL := 21214,
	ILLEGALPARAMETER_MOVEDIRREL := 21215,
	NOVALIDVELOCITY_MANMODE := 21216,
	NOVALIDACCELERATION_MANMODE := 21217,
	NOVALIDDECELERATION_MANMODE := 21218,
	NOVALIDJERK_MANMODE := 21219,
	MANUALMODEILLEGALPARAMETER := 21220,
	KINEMATICILLEGALPARAMETER := 21221,
	AXESGROUPINERRORSTOP := 21222,
	TOOLINUSE := 21223,
	INVALIDTOOL := 21224,
	AXESGROUPINMOVEMENT := 21225,
	INVALIDCOORDSYSTEM := 21226,
	AXISEXTERNALENABLED := 21227,
	UNSUPPORTEDCOORDSYSTEM := 21228,
	REALAXISNOTREADY := 21229,
	INVALIDAXESGROUPSTATE := 21230,
	REALAXISOUTSIDEWORKINGRANGE := 21231,
	SINGULARPOSITION := 21232,
	L_MC4P_INTERNALERROR := 21233,
	AXESGROUPEXTERNALSTOPPING := 21234,
	RESETAXESGROUPERRORFAILED := 21237,
	ILLEGALTEACHPOSITION := 21238,
	NOTENOUGHMEMORYPATHDATALIST := 21239,
	NOVALIDROTATIONVELOCITY_MOVECIRCABS := 21240,
	NOVALIDROTATIONACCELERATION_MOVECIRCABS := 21241,
	NOVALIDROTATIONJERK_MOVECIRCABS := 21242,
	NOVALIDROTATIONVELOCITY_MOVECIRCREL := 21243,
	NOVALIDROTATIONACCELERATION_MOVECIRCREL := 21244,
	NOVALIDROTATIONJERK_MOVECIRCREL := 21245,
	NOVALIDROTATIONVELOCITY_MOVELINABS := 21246,
	NOVALIDROTATIONACCELERATION_MOVELINABS := 21247,
	NOVALIDROTATIONJERK_MOVELINABS := 21248,
	NOVALIDROTATIONVELOCITY_MOVELINREL := 21249,
	NOVALIDROTATIONACCELERATION_MOVELINREL := 21250,
	NOVALIDROTATIONJERK_MOVELINREL := 21251,
	PATHLIMITVIOLATION_MOVELINABS := 21252,
	PATHLIMITVIOLATION_MOVELINREL := 21253,
	PATHLIMITVIOLATION_MOVECIRCABS := 21254,
	PATHLIMITVIOLATION_MOVECIRCREL := 21255,
	PATHLIMITVIOLATION_MOVEDIRABS := 21256,
	PATHLIMITVIOLATION_MOVEDIRREL := 21257,
	AXISGROUPNOTHOMED := 21258,
	MAINAXISTYPEMODULONOTALLOWED := 21259,
	AXISTYPEMODULONOTALLOWED := 21260,
	AXISLIMITVIOLATIONREALAXIS1VELOCITY := 21261,
	AXISLIMITVIOLATIONREALAXIS2VELOCITY := 21262,
	AXISLIMITVIOLATIONREALAXIS3VELOCITY := 21263,
	AXISLIMITVIOLATIONREALAXIS4VELOCITY := 21264,
	AXISLIMITVIOLATIONREALAXIS5VELOCITY := 21265,
	AXISLIMITVIOLATIONREALAXIS6VELOCITY := 21266,
	AXISLIMITVIOLATIONREALAXIS1ACCELERATION := 21267,
	AXISLIMITVIOLATIONREALAXIS2ACCELERATION := 21268,
	AXISLIMITVIOLATIONREALAXIS3ACCELERATION := 21269,
	AXISLIMITVIOLATIONREALAXIS4ACCELERATION := 21270,
	AXISLIMITVIOLATIONREALAXIS5ACCELERATION := 21271,
	AXISLIMITVIOLATIONREALAXIS6ACCELERATION := 21272,
	AUXAXISSEQUENCEINVALID := 21273,
	AUXAXISNOTALLOWED := 21274,
	ILLEGALTRACKINGPARAMETER := 21275,
	SYNCHRONISATIONERROR := 21276,
	PCSINUSE := 21277,
	TRACKINGFBNOTCALLED := 21278,
	MASTERAXISNOTREADY := 21279,
	MOVEDIRECTNOTALLOWED := 21280,
	AUXAXISNOVALIDVELOCITY := 21281,
	AUXAXISNOVALIDACCELERATION := 21282,
	AUXAXISNOVALIDJERK := 21283,
	MAINAXISNOTCONNECTED := 21284,
	REALAXISNOTCONNECTED := 21285,
	AXESGROUPNOTINITIALIZED := 21286,
	DISABLEDBYPARAMETERTRANSFER := 21287,
	REALAXIS1_ALREADYINUSE := 21288,
	REALAXIS2_ALREADYINUSE := 21289,
	REALAXIS3_ALREADYINUSE := 21290,
	REALAXIS4_ALREADYINUSE := 21291,
	REALAXIS5_ALREADYINUSE := 21292,
	REALAXIS6_ALREADYINUSE := 21293,
	AUXAXIS1_ALREADYINUSE := 21294,
	AUXAXIS2_ALREADYINUSE := 21295,
	AUXAXIS3_ALREADYINUSE := 21296,
	AUXAXIS4_ALREADYINUSE := 21297,
	AUXAXIS5_ALREADYINUSE := 21298,
	AUXAXIS6_ALREADYINUSE := 21299,
	NOVALIDTRANSITIONMODE_MOVECIRCABS := 21300,
	NOVALIDTRANSITIONMODE_MOVECIRCREL := 21301,
	NOVALIDTRANSITIONMODE_MOVELINABS := 21302,
	NOVALIDTRANSITIONMODE_MOVELINREL := 21303,
	NOVALIDTRANSITIONMODE_MOVEDIRABS := 21304,
	NOVALIDTRANSITIONMODE_MOVEDIRREL := 21305,
	NOAXISFORHOMINGSELECTED := 21306,
	INVALIDTARGETORIENTATION := 21307,
	NOKINTRANSFORMATIONAVAILABLE := 21308,
	AXESGROUPNOTSUPPORTED := 21309,
	AXESGROUPNOTDISABLED := 21310,
	AXESGROUPINITFAILED := 21311,
	KINTRANSFORMATIONINUSE := 21312,
	MAXNUMREVOLUTIONSREACHED := 21313,
	PCSCHANGEDDURINGMOTION := 21314,
	CONCURRENTREQUESTMANUALMODE := 21315,
	PATHREFCOMMANDNOTSUPPORTED := 21316,
	PATHREFSYNTAXERROR := 21317,
	PATHREFGCOMMANDNOTSUPPORTED := 21318,
	PATHREFMCOMMANDNOTSUPPORTED := 21319,
	PATHREFINVALIDCOMENTSYNTAX := 21320,
	FILEACCESSTIMEOUT := 21321,
	INVALIDPATHREF := 21322,
	INVALIDPATHFILE := 21323,
	IJKCOMMANDMISSING := 21324,
	INVALIDCIRCCOMMAND := 21325,
	DYNAMICCHANGEOFPATHREFNOTALLOWED := 21327,
	CONCURRENTMFUNCTION := 21328,
	INVALIDMSTARTRADIUSGTSEMIMAJORAXISSTARTRADIUSLTSEMIMINORAXISTARGETRADIUSGTSEMIMAJORAXISFUNCTION := 21329,
	STARTRADIUSGTSEMIMAJORAXIS := 21330,
	STARTRADIUSLTSEMIMINORAXIS := 21331,
	TARGETRADIUSGTSEMIMAJORAXIS := 21332,
	TARGETRADIUSLTSEMIMINORAXIS := 21333,
	SEMIMINORAXISGTSEMIMAJORAXIS := 21334,
	SEMIMINORAXISLE0 := 21335,
	SEMIMAJORAXISLE0 := 21336,
	TARGETNOTONELLIPSE := 21337,
	INVALIDTRAVERSINGRANGECOMBINATION := 21338,
	INVALIDCOORDINATESYSTEMORIENTATION := 21339,
	INVALIDTOOLSYSTEMORIENTATION := 21340,
	TARGETNOTONCIRC := 21341,
	EXECUTIONLOCKEDBYMOVEPATH := 21342,
	NOVALIDVELOCITY_MOVESPLINE := 21343,
	NOVALIDACCELERATION_MOVESPLINE := 21344,
	NOVALIDDECELERATION_MOVESPLINE := 21345,
	NOVALIDJERK_MOVESPLINE := 21346,
	NOVALIDTRANSITIONPARAMETER_MOVESPLINE := 21347,
	NOVALIDTRANSITIONMODE_MOVESPLINE := 21348,
	POSITIONOUTSIDESWLIMITSMAINAXISX_MOVESPLINE := 21349,
	POSITIONOUTSIDESWLIMITSMAINAXISY_MOVESPLINE := 21350,
	POSITIONOUTSIDESWLIMITSMAINAXISZ_MOVESPLINE := 21351,
	POSITIONOUTSIDESWLIMITSMAINAXISA_MOVESPLINE := 21352,
	POSITIONOUTSIDESWLIMITSMAINAXISB_MOVESPLINE := 21353,
	POSITIONOUTSIDESWLIMITSMAINAXISC_MOVESPLINE := 21354,
	NOVALIDROTATIONVELOCITY_MOVESPLINE := 21355,
	NOVALIDROTATIONACCELERATION_MOVESPLINE := 21356,
	NOVALIDROTATIONJERK_MOVESPLINE := 21357,
	NOINTERMEDIATEPOINTS_MOVESPLINE := 21358,
	PATHLIMITVIOLATION_MOVESPLINE := 21359,
	NOVALIDINTERMEDIATEPOINTLOCATION := 21360,
	POSITIONOUTSIDESWLIMITSREALAXIS1_MOVESPLINE := 21361,
	POSITIONOUTSIDESWLIMITSREALAXIS2_MOVESPLINE := 21362,
	POSITIONOUTSIDESWLIMITSREALAXIS3_MOVESPLINE := 21363,
	POSITIONOUTSIDESWLIMITSREALAXIS4_MOVESPLINE := 21364,
	POSITIONOUTSIDESWLIMITSREALAXIS5_MOVESPLINE := 21365,
	POSITIONOUTSIDESWLIMITSREALAXIS6_MOVESPLINE := 21366,
	POSITIONOUTSIDESWLIMITSAUXAXIS1_MOVESPLINE := 21367,
	POSITIONOUTSIDESWLIMITSAUXAXIS2_MOVESPLINE := 21368,
	POSITIONOUTSIDESWLIMITSAUXAXIS3_MOVESPLINE := 21369,
	POSITIONOUTSIDESWLIMITSAUXAXIS4_MOVESPLINE := 21370,
	POSITIONOUTSIDESWLIMITSAUXAXIS5_MOVESPLINE := 21371,
	POSITIONOUTSIDESWLIMITSAUXAXIS6_MOVESPLINE := 21372,
	POSITIONTRANSFORMATIONERROR_MOVESPLINE := 21373,
	POSITIONOUTSIDESWLIMITSPASSIVEJOINTS_MOVESPLINE := 21374,
	POSITIONSINGULARPOS_MOVESPLINE := 21375,
	CONCURRENTTORQUEPRECONTROL := 21376,
	INVALIDORIENTATIONMODE := 21377,
	CONCURRENTAXESGROUPBASICCONTROL := 21378,
	PARAMETERLIMITSNOTSUFFICIENT := 21379,
	SETVALUEMANIPULATIONNOTSUPPORTED := 21380,
	MINPOSGTMAXPOS := 21381,
	DYNAMICPARAMETERNOTPLAUSIBLE := 21382,
	CONVERGENCENOTSUFFICIENT := 21383,
	IDENTIFICATIONNOTDONE := 21384,
	INVALIDOVERRIDEFORIDENTIFICATION := 21385,
	PHASINGNOTALLOWED := 22000,
	INVALIDCAMREF := 22010,
	INVALIDCAMTYPE := 22011,
	INVALIDCAMDATA := 22012,
	INVALIDDATACOUNT := 22013,
	DATACOUNTTOOSMALL := 22014,
	INVALIDLAWOFMOTION := 22015,
	INVALIDINPUTDATA := 22016,
	MASTEROUTOFCAM := 22025,
	INVALIDVELACC_OFFSETSCALING := 22026,
	INVALIDCAMTABLE := 22027,
	INVALIDSTARTORENDPOSOFCAM := 22028,
	INVALIDSCALINGFACTOR := 22029,
	RAMPINERROR := 22030,
	NOTALLOWEDMOVEMENTBYMASTER := 22035,
	CLUTCHISREVERSING := 22036,
	INVALIDDEFAULTJERK := 22037,
	INVALIDOPENINSTANTDEC := 22038,
	INVALIDREVERSE := 22039,
	FILENOTFOUND := 22050,
	INVALIDFILE := 22051,
	INVALIDCHECKCRC := 22052,
	INVALIDDATASIZE := 22053,
	INVALIDTAPPETREF := 22060,
	INVALIDTAPPETDATA := 22061,
	INVALIDTAPPETTYPE := 22062,
	INVALIDTIMINGTAPPET := 22063,
	INVALIDPOSSELECTIONTAPPET := 22064,
	DYNAMISATIONERROR := 22065,
	XCYCLELENGTHINVALID_LINEARCOUPLING := 22082,
	YCYCLELENGTHINVALID_LINEARCOUPLING := 22083,
	POSININVALID_LINEARCOUPLING := 22084,
	INVALIDTAPPETSCOUNT := 22085,
	RESETPHASINGNOTALLOWED := 22086
);
END_TYPE

(* ---- OEEWEEKDAY.dut ---- *)
TYPE OEEWEEKDAY :
(
	SUNDAY := 0,
	MONDAY := 1,
	TUSEDAY := 2,
	WEDNESDAY := 3,
	THURSDAY := 4,
	FRIDAY := 5,
	SATURDAY := 6
);
END_TYPE

(* ---- SCAXISPOSCOUNT.dut ---- *)
TYPE SCAXISPOSCOUNT :
STRUCT
	LRAXISPOSINT : LREAL;
	LRAXISPOSCOUNTINT : LREAL;
	LRLASTAXISPOS : LREAL;
	LRDIFFAXISPOS : LREAL;
END_STRUCT
END_TYPE

(* ---- SCCATEGORYSTRUCT.dut ---- *)
TYPE SCCATEGORYSTRUCT :
STRUCT
	ASSTR : ARRAY [0..uiNoOfDowntimeCategories] OF STRING(55);
	AXERROR : ARRAY [0..uiNoOfDowntimeCategories] OF BOOL;
END_STRUCT
END_TYPE

(* ---- SCCLOUDDATA.dut ---- *)
TYPE SCCLOUDDATA :
STRUCT
	XSTATECHANGEPROLONGED : BOOL;
	ITRIGGER : INT;
	XSHIFTDATAPROLONGED : BOOL;
	SEVENT : STRING(255);
	SSHIFTOEEKPIS : STRING(255);
	SPRODUCTOEEKPIS : STRING(255);
	SSTATIONNAME : STRING;
END_STRUCT
END_TYPE

(* ---- SCDATETIMEMONITORING.dut ---- *)
TYPE SCDATETIMEMONITORING :
STRUCT
	DTLASTMACHINEDATETIME : DATE_AND_TIME;
	DTLASTLINEDATETIME : DATE_AND_TIME;
	TDATETIMEDEVIATION : TIME;
	TDATETIMECONNECTION : TIME;
END_STRUCT
END_TYPE

(* ---- SCERRORDATA.dut ---- *)
TYPE SCERRORDATA :
STRUCT
	XFIRSTERRORACTIVE : BOOL;
	XISWARNINGINFO : BOOL;
	IPRIORITY : INT;
	DWERRORNUMBER : DWORD;
END_STRUCT
END_TYPE

(* ---- SCERRORDATA_BASE.dut ---- *)
TYPE SCERRORDATA_BASE :
STRUCT
	SERRDESC : STRING;
	SCATEGORYDESC : STRING(55);
	DWERRORCATEGORY : DWORD;
	PRODUCTIONEVENTMODE : INT;
	XCATEGORYERROR : BOOL;
END_STRUCT
END_TYPE

(* ---- SCEXECUTETIME.dut ---- *)
TYPE SCEXECUTETIME :
STRUCT
	SFBSTR : STRING;
	LRLASTTIME : LREAL;
	LRTIMEAVEARAGE : LREAL;
	LRMAXTIME : LREAL;
	LRCOUNT : LREAL;
	LRTIMESUMCOUNT : LREAL;
	LRLASTTIMEAVEARAGE : LREAL;
END_STRUCT
END_TYPE

(* ---- SCEXECUTETIMEARRAY.dut ---- *)
TYPE SCEXECUTETIMEARRAY :
STRUCT
	AEXECUTION : ARRAY [1..15] OF scExecuteTime;
END_STRUCT
END_TYPE

(* ---- SCLINEKPIS.dut ---- *)
TYPE SCLINEKPIS :
STRUCT
	ILINEID : INT;
	SLINEID : STRING;
	SDATETIME : STRING;
	SSHIFTNAME : STRING;
	ROEERT : REAL;
	RTEEP : REAL;
	RAVAILABILITY : REAL;
	RPERFORMANCE : REAL;
	RQUALITY : REAL;
	LRQUANTITYOK : LREAL;
	LRQUANTITYNOK : LREAL;
	LRQUANTITYOKTOTAL : LREAL;
	LRQUANTITYNOKTOTAL : LREAL;
	DIACTUALRUNTIME : DINT;
	DIDOWNTIME : DINT;
	DIORGDOWNTIME : DINT;
	DINONPRODUCTIVETIME : DINT;
	DIACTUALRUNTIMETOTAL : DINT;
	DIDOWNTIMETOTAL : DINT;
	DIORGDOWNTIMETOTAL : DINT;
	DINONPRODUCTIVETIMETOTAL : DINT;
	XSHIFTDATAPROLONGED : BOOL;
END_STRUCT
END_TYPE

(* ---- SCLINESTATUS.dut ---- *)
TYPE SCLINESTATUS :
STRUCT
	XALLMACHINECONNECTED : BOOL;
	XALLMACHINEDATETIMEINSYNCH : BOOL;
	XALLMACHINEACTIVE : BOOL;
	XALLMACHINEACTIVEOEECALC : BOOL;
	INOCONNECTEDMACHINE : INT;
	INODATETIMEINSYNCH : INT;
	INOMACHINEACTIVE : INT;
	INOMACHINEACTIVEOEECALC : INT;
	IINDEXFIRSTMACHINENOTCONNECTED : INT;
	IINDEXFIRSTMACHINENOTDATETIMEINSYNCH : INT;
	IINDEXFIRSTMACHINENOTACTIVE : INT;
	SNAMEFIRSTMACHINENOTCONNECTED : STRING;
	SNAMEFIRSTMACHINENOTDATETIMEINSYNCH : STRING;
	SNAMEFIRSTMACHINENOTACTIVE : STRING;
	SIPADDRESSFIRSTMACHINENOTCONNECTED : STRING;
	SIPADDRESSFIRSTMACHINENOTDATETIMEINSYNCH : STRING;
	SIPADDRESSFIRSTMACHINENOTACTIVE : STRING;
END_STRUCT
END_TYPE

(* ---- SCMACHINEDATA_NVL.dut ---- *)
TYPE SCMACHINEDATA_NVL :
STRUCT
	SMACHINENAME : STRING;
	SIPADDRESS : STRING;
	XCONNECTED : BOOL;
	XDATETIMEINSYNCH : BOOL;
	XACTIVEOEECALC : BOOL;
	SCDTMONITOR : scDateTimeMonitoring;
	ROEE_WEIGHT : REAL;
END_STRUCT
END_TYPE

(* ---- SCMACHINEOFFMODE.dut ---- *)
TYPE SCMACHINEOFFMODE :
STRUCT
	IPRODUCTIONMODE : INT := 0;
	IDOWNTIMECATEGORY : INT := 0;
	UDIDOWNTIMEREASON : UINT := 0;
	SINTERVAL : STRING := '';
	ASDOWNTIMESTR : STRING := '';
	SREASONCODE : STRING := '';
END_STRUCT
END_TYPE

(* ---- SCMACHINESHIFTACTIVE.dut ---- *)
TYPE SCMACHINESHIFTACTIVE :
STRUCT
	DTACTIVEDURINGACTUALSHIFT : DATE_AND_TIME;
	XACTIVEDURINGACTUALSHIFT : BOOL;
END_STRUCT
END_TYPE

(* ---- SCOEE_NVL.dut ---- *)
TYPE SCOEE_NVL :
STRUCT
	SDATETIME : STRING;
	SCPERFORMANCEKPI : scPerformance_base;
	SCPERFORMANCEADDS : scOEE_Substructurs;
	SCRR : scRunRate;
	SCCLOUDDATA : scCloudData;
	XACTIVE : BOOL;
END_STRUCT
END_TYPE

(* ---- SCOEE_SUBSTRUCTURS.dut ---- *)
TYPE SCOEE_SUBSTRUCTURS :
STRUCT
	LRACTUALTHROUGHPUT_HR : LREAL;
	LRTARGETTHROUGHPUT_HR : LREAL;
	SINTERVAL : STRING;
	SDOWNTIMESTR : STRING;
	SREASONCODE : STRING;
	RSETSPEEDVALUE : REAL;
	RSETSPEEDPERCENT : REAL;
	ITRIGGER : INT;
	DIACTUALPLANNEDPRODUCTION : DINT;
	DIACTUALRUNTIME : DINT;
	DIDOWNTIME : DINT;
	DIORGDOWNTIME : DINT;
	DINONPRODUCTIVETIME : DINT;
	DISTATERUNTIME : DINT;
	DISTATETOTALTIME : DINT;
	ITRIGGER_SETTINGS : INT;
	XSHIFTCHANGESTOREEVENT : BOOL;
END_STRUCT
END_TYPE

(* ---- SCPRODUCTIONMODE.dut ---- *)
TYPE SCPRODUCTIONMODE :
STRUCT
	ASMODE : ARRAY [0..uiNoOfProductionModes] OF STRING;
	SMODECOLOURCODE : ARRAY [0..uiNoOfProductionModes] OF STRING(6);
END_STRUCT
END_TYPE

(* ---- SCREF_NVL.dut ---- *)
TYPE SCREF_NVL :
STRUCT
	SCOEE_NVL : REFERENCE TO scOEE_NVL;
END_STRUCT
END_TYPE

(* ---- SCSHIFTNAME.dut ---- *)
TYPE SCSHIFTNAME :
STRUCT
	ESETWEEKDAY : RTCLK.WEEKDAY;
	SSETSHIFTNAME : STRING;
	XUSEWEEKDAY : BOOL;
END_STRUCT
END_TYPE

(* ---- SCSIMULATIONDOWNTIMES.dut ---- *)
TYPE SCSIMULATIONDOWNTIMES :
STRUCT
	UIMAXSIMULATIONEVENTS : UINT := 13;
	SCRT : RT_Downtime := STRUCT(para := [STRUCT(DowntimeCode := 5, ProductionMode := 2, ReasonCode := 16#3C000001, sReasonCodeStr := 'Stopping for long'), STRUCT(DowntimeCode := 6, ProductionMode := 9, ReasonCode := 16#3C000002, sReasonCodeStr := 'Drive-24V Supply'), STRUCT(DowntimeCode := 7, ProductionMode := 9, ReasonCode := 16#3C000008, sReasonCodeStr := 'Power supply error'), STRUCT(DowntimeCode := 3, ProductionMode := 9, ReasonCode := 16#3C000004, sReasonCodeStr := 'Emergency Stop'), STRUCT(DowntimeCode := 5, ProductionMode := 2, ReasonCode := 16#3C000005, sReasonCodeStr := 'Line Speed 0'), STRUCT(DowntimeCode := 5, ProductionMode := 6, ReasonCode := 16#3C000006, sReasonCodeStr := 'Line Speed < 100'), STRUCT(DowntimeCode := 1, ProductionMode := 5, ReasonCode := 16#3C00000C, sReasonCodeStr := 'No Parts'), STRUCT(DowntimeCode := 3, ProductionMode := 9, ReasonCode := 16#3C000007, sReasonCodeStr := 'Safety light curtain interrupted'), STRUCT(DowntimeCode := 6, ProductionMode := 9, ReasonCode := 16#3C00000D, sReasonCodeStr := 'Drive over-temperature'), STRUCT(DowntimeCode := 11, ProductionMode := 6, ReasonCode := 16#3C00000A, sReasonCodeStr := 'Rotation Limit detected'), STRUCT(DowntimeCode := 12, ProductionMode := 10, ReasonCode := 16#0, sReasonCodeStr := ''), STRUCT(DowntimeCode := 12, ProductionMode := 10, ReasonCode := 16#3C00000F, sReasonCodeStr := 'Time exceeded'), STRUCT(DowntimeCode := 5, ProductionMode := 6, ReasonCode := 16#3C00000E, sReasonCodeStr := 'Recipe change'), STRUCT(DowntimeCode := 0, ProductionMode := 0, ReasonCode := 16#0, sReasonCodeStr := ''), STRUCT(DowntimeCode := 0, ProductionMode := 0, ReasonCode := 16#0, sReasonCodeStr := ''), STRUCT(DowntimeCode := 0, ProductionMode := 0, ReasonCode := 16#0, sReasonCodeStr := ''), STRUCT(DowntimeCode := 0, ProductionMode := 0, ReasonCode := 16#0, sReasonCodeStr := ''), STRUCT(DowntimeCode := 0, ProductionMode := 0, ReasonCode := 16#0, sReasonCodeStr := ''), STRUCT(DowntimeCode := 0, ProductionMode := 0, ReasonCode := 16#0, sReasonCodeStr := ''), STRUCT(DowntimeCode := 0, ProductionMode := 0, ReasonCode := 16#0, sReasonCodeStr := '')]);
	SCRECIPE : ARRAY [0..1] OF scProduct_base := [STRUCT(rTechnicalCycleTime := 1.5, rProductTarget := 15480, diTypeID := 1, sTypeName := 'Biscuit Box', iUnitProductID := 1, sUnitProduct := 'Boxes', iUnitSpeedID := 1, sUnitSpeed := 'Boxes/min.'), STRUCT(rTechnicalCycleTime := 1.25, rProductTarget := 18576, diTypeID := 2, sTypeName := 'Chocolate Box', iUnitProductID := 1, sUnitProduct := 'Boxes', iUnitSpeedID := 1, sUnitSpeed := 'Boxes/min.')];
END_STRUCT
END_TYPE

(* ---- SCSIMULATIONMODES.dut ---- *)
TYPE SCSIMULATIONMODES :
STRUCT
	DOWNTIMEACTIVE1 : INT := 9;
	DOWNTIMEACTIVE2 : INT;
	ORGDOWNTIMEACTIVE1 : INT := 2;
	ORGDOWNTIMEACTIVE2 : INT := 5;
	ORGDOWNTIMEACTIVE3 : INT := 10;
END_STRUCT
END_TYPE

(* ---- GVL_AXISSIM.gvl ---- *)
VAR_GLOBAL
	FEEDERAXIS : AXIS_REF_SIM := STRUCT(eTraversingRange := 1, lrCycleLength := 1000.0, lrFeedConstant := 1000.0, dwGearNumerator := 100, dwGearDenominator := 1, eMctrlMode := 0, wNoOfHTLPeriods := 128);
END_VAR

(* ---- GVL_VALIDATIONTEST.gvl ---- *)
VAR_GLOBAL
	SCEXECUTETIMEARRAY : scExecuteTimeArray;
	SCMACHINEDATA_BASE : scMachineData_base;
	SCPERFORMANCE_BASE : scPerformance_base;
	ULISTART : ULINT;
	ULIEND : ULINT;
	XPRODUCTIONACTIVE : BOOL := TRUE;
	FBMACHINEPERFORMANCE_BASE : L_OEEA_MachinePerformance_Base;
	FBDOWNTIME_BASE : L_OEEA_Downtime_base;
	FBSHIFTOEEHISTORYALL : L_OEEA_ShiftOEEHistory;
	FBSHIFTOEEHISTORY_BASE : L_OEEA_ShiftOEEHistory_Base;
	FBSHIFTDOWNTIMEHISTORY_BASE : L_OEEA_ShiftDowntimeHistory_base;
	SCPDINTERNAL_BASE : scInternalVar;
	SCPDSHIFTDAYINDEX : scPDShiftData;
	SCPDINTERNALDOWNTIME_BASE : scInternalDownVar;
	SCDOWNTIME_BASE : scDowntime_base;
	SCSHIFTDOWNTIMEHISTORY_BASE : ARRAY [1..3] OF scDowntime_base;
	SCSHIFTHISTORYALL : ARRAY [1..3] OF scPerformance;
	SCPDSHIFTHISTORY_BASE : scVisuShiftHistory_base;
	SCPDPRODUCTIONDATA : scInternalProductionData;
	SCSHIFTVALUES : scCurrentShiftValues;
END_VAR

(* ---- LINE_OEE_GVL_VAR.gvl ---- *)
VAR_GLOBAL
	UINOOFMACHINES : UINT := 60;
	UINOOFHISTORICALWEEKS : UINT := 4;
END_VAR

(* ---- VERSIONCONSTANTS.gvl ---- *)
VAR_GLOBAL
	GC_BYAMOUNTOFGENERALDATA : BYTE := 50;
	GC_BYAMOUNTDOWNTIMEERRORS : BYTE := 10;
	GC_IFILTERSAMPLES : INT := 20;
END_VAR

(* ---- CALENDAR_WEEK.pou ---- *)
FUNCTION CALENDAR_WEEK : UINT
VAR_INPUT
	DTEXTDT : DATE_AND_TIME;
END_VAR
END_FUNCTION

(* ---- EXECUTIONTIME.pou ---- *)
FUNCTION EXECUTIONTIME : BOOL
VAR_INPUT
	SFBSTR : STRING;
	ULISTART : ULINT;
	ULIEND : ULINT;
END_VAR
VAR_IN_OUT
	AEXECUTION : scExecuteTime;
END_VAR
END_FUNCTION

(* ---- L_OEEA_CUSTOMIZABLE_COPYSTRUCT.pou ---- *)
FUNCTION L_OEEA_CUSTOMIZABLE_COPYSTRUCT : BOOL
VAR_INPUT
	PBYSOURCE : POINTER TO BYTE;
	PBYTARGET : POINTER TO BYTE;
	UISIZESOURCE : UINT;
	UISIZETARGET : UINT;
END_VAR
END_FUNCTION

(* ---- LRAXISPOSCOUNT.pou ---- *)
FUNCTION LRAXISPOSCOUNT : LREAL
VAR_INPUT
	LRAXISPOS : LREAL;
END_VAR
VAR_IN_OUT
	SCAXISPOSCOUNT : scAxisPosCount;
END_VAR
END_FUNCTION

(* ---- GLOBALTEXTLIST.pou ---- *)
FUNCTION_BLOCK GLOBALTEXTLIST
VAR
	M_TEXTLISTFILE : STRING(255);
	_STNAMESPACE : STRING;
END_VAR
END_FUNCTION_BLOCK

(* ---- IMAGEPOOL_AXIS_REF_SIM.pou ---- *)
FUNCTION_BLOCK IMAGEPOOL_AXIS_REF_SIM
VAR
	M_STNAMESPACE : STRING(80);
	M_STHELPVARID : STRING;
	M_STHELPVARPATH : STRING(255);
	M_STHELP : STRING;
	M_REGISTERIMAGES : BOOL := TRUE;
END_VAR
END_FUNCTION_BLOCK

METHOD FB_INIT : BOOL
VAR_INPUT
	BINITRETAINS : BOOL;
	BINCOPYCODE : BOOL;
END_VAR
END_METHOD

METHOD FB_REINIT : BOOL
END_METHOD

METHOD FB_EXIT : BOOL
VAR_INPUT
	BINCOPYCODE : BOOL;
END_VAR
END_METHOD

(* ---- L_MC1A_BASICACTUATINGSPEED.pou ---- *)
FUNCTION_BLOCK L_MC1A_BASICACTUATINGSPEED
VAR_INPUT
	XREGULATORON : BOOL;
	XRESETERROR : BOOL;
	XSETDRIVEQSP : BOOL;
	XENABLESETVEL : BOOL;
	XINVERTDIRECTION : BOOL;
	LRSETVEL : LREAL := 300.0;
	LRSETACC : LREAL := 100.0;
	LRSETDEC : LREAL := 100.0;
END_VAR
VAR_OUTPUT
	XERROR : BOOL;
	XBUSY : BOOL;
	EERRORID : L_IE1A_ErrorID;
	XCOMMUNICATIONOK : BOOL;
	XAXISREADY : BOOL;
	XAXISENABLED : BOOL;
	XDRIVEWARNING : BOOL;
	XDRIVEERROR : BOOL;
	DWDRIVEERRORID : DWORD;
	XDRIVEQSPACTIVE : BOOL;
	LRACTVEL : LREAL;
	XDIRECTIONPOSITIVE : BOOL;
	XDIRECTIONNEGATIVE : BOOL;
	WDIGITALINPUTS : WORD;
END_VAR
VAR_IN_OUT
	AXIS : AXIS_REF_SIM;
END_VAR
VAR
	L_TB1A_PT1FILTER1 : L_TB1A_PT1Filter := STRUCT(lrFilterTime := 0.02);
	L_MC1A_INTEGRATEAXIS1 : L_MC1A_IntegrateAxis;
	L_MC1A_DIFFERENTIATE2 : L_MC1A_Differentiate;
	L_MC1A_CONVX1 : L_MC1A_ConvX := STRUCT(diDenom := 1000000000);
	L_MC1A_CONVX2 : L_MC1A_ConvX;
	R_TRIG3 : R_TRIG;
	TON0 : TON := STRUCT(IN := TRUE, PT := TIME#1m0s0ms);
	TON1 : TON;
	TP1 : TP;
	X1STCYCLE : BOOL := TRUE;
	BYINITCOUNTER : BYTE;
	LRTASKCYCLETIME : LREAL;
	DITASKCYCLETIME : DINT;
	XINIT : BOOL := TRUE;
	LRACTVEL_INTERNAL : LREAL;
	LRREVPERSEC : LREAL;
	LITMP1 : LINT;
	LITMP2 : LINT;
	LITMP3 : LINT;
	LITMP6 : LINT;
	LITMP7 : LINT;
	RRANDOMNUMBER : REAL;
	RTMP : REAL;
	RHEATSINKTEMPINT : REAL;
	RHEATSINKFILTERTIME : REAL := 73.7;
	RIXTLOADINT : REAL;
	RIXTLOADFILTERTIME : REAL := 43.3;
	RIXT2LOADINT : REAL;
	RIXT2LOADFILTERTIME : REAL := 37.3;
	LROPERATIONTIME : LREAL;
	LROPERATIONTIMECU : LREAL;
	LRMODULOCYCLELENGTH_INTERNAL : LREAL;
	DIMODULOCYCLELENGTH_INTERNAL : DINT;
	LRPOSTOUNITFACTOR : LREAL;
	LRTMPEE : LREAL;
	DWMODULOCYCLERESIDUAL : DWORD;
	DIHALFMODULOCYCLELENGTH : DINT;
	DWRESIDUAL : DWORD;
	DIACTPOS : DINT;
	DIACTPOSOLD : DINT;
	XRESADDACTCYCLE : BOOL;
	XRESSUBACTCYCLE : BOOL;
	DWHTLCOUNTERVALUE_INTERNAL : DWORD;
	DIDELTAPOS : DINT;
	DIINPUTOLD : DINT;
	DITMPEE : DINT;
END_VAR
END_FUNCTION_BLOCK

METHOD METH_RAMPGENERATOR : LREAL
VAR_INPUT
	LRSETVEL : LREAL;
	LRSETACC : LREAL;
	LRSETDEC : LREAL;
	LRACTVEL : LREAL;
	XLOADSTARTVEL : BOOL;
	LRSTARTVEL : LREAL;
END_VAR
END_METHOD

METHOD ACT_SDOEMULATION
END_METHOD

METHOD METH_RANDOM : REAL
VAR_INPUT
	RRANDOMNUMBER : REAL;
END_VAR
END_METHOD

(* ---- L_MC1A_CONVX.pou ---- *)
FUNCTION_BLOCK L_MC1A_CONVX
VAR_INPUT
	DIIN : DINT;
	DINUM : DINT := 1;
	DIDENOM : DINT := 1;
END_VAR
VAR_OUTPUT
	DIOUT : DINT;
	XLIMIT : BOOL;
END_VAR
VAR
	LIOUT : LINT;
	LIREMAINDER : LINT;
	LITMP : LINT;
	LIDENOMINATOR : LINT;
END_VAR
END_FUNCTION_BLOCK

(* ---- L_MC1A_DIFFERENTIATE.pou ---- *)
FUNCTION_BLOCK L_MC1A_DIFFERENTIATE
VAR_INPUT
	LRPOSITIONIN : LREAL;
	ETRAVERSINGRANGE : WORD;
	LRCYCLELENGTH : LREAL := 360.0;
END_VAR
VAR_OUTPUT
	LRVELOCITYOUT : LREAL;
	XERROR : BOOL;
END_VAR
VAR
	TON0 : TON := STRUCT(IN := TRUE, PT := TIME#1m0s0ms);
	X1STCYCLE : BOOL := TRUE;
	BYINITCOUNTER : BYTE;
	LRTASKCYCLETIME : LREAL;
	LRCYCLELENGTHINTERNAL : LREAL;
	LRPOSITIONINLIMITED : LREAL;
	LRPOSITIONINLIMITEDOLD : LREAL;
END_VAR
END_FUNCTION_BLOCK

METHOD METH_SHORTESTWAY : LREAL
VAR_INPUT
	LRSETPOS : LREAL;
	LRACTPOS : LREAL;
	LRCYCLELENGTH : LREAL;
END_VAR
END_METHOD

(* ---- L_MC1A_INTEGRATEAXIS.pou ---- *)
FUNCTION_BLOCK L_MC1A_INTEGRATEAXIS
VAR_INPUT
	LRVELIN : LREAL;
	XLOADSTARTPOSITION : BOOL;
	LRSTARTPOSITION : LREAL;
	LRCYCLELENGTH : LREAL;
END_VAR
VAR_OUTPUT
	LRPOSOUT : LREAL;
	LRVELOUT : LREAL;
	XZEROCW : BOOL;
	XZEROCCW : BOOL;
	XZERO : BOOL;
END_VAR
VAR
	TON0 : TON := STRUCT(IN := TRUE, PT := TIME#1m0s0ms);
	X1STCYCLE : BOOL := TRUE;
	BYINITCOUNTER : BYTE;
	LRTASKCYCLETIME : LREAL;
	LRPOSOUT_OLD : LREAL;
END_VAR
END_FUNCTION_BLOCK

METHOD METH_ADDOFFSETCYCLIC : LREAL
VAR_INPUT
	LRSETPOS : LREAL;
	LRSETOFFSET : LREAL;
	LRCYCLELENGTH : LREAL;
END_VAR
END_METHOD

(* ---- L_OEEA_BASE_FBS.pou ---- *)
FUNCTION_BLOCK L_OEEA_BASE_FBS EXTENDS L_OEEA_FBs_COMMON
VAR_IN_OUT
	SCMACHINEDATA_BASE : scMachineData_base;
	SCPERFORMANCE_BASE : scPerformance_base;
	SCDOWNTIME_BASE : scDowntime_base;
END_VAR
VAR
	FBMACHINEPERFORMANCE : L_OEEA_MachinePerformance_Base;
	SCMACHINEDATA : scMachineData;
	FBDOWNTIME : L_OEEA_Downtime_Base;
	SCDOWNTIME : scDowntime;
END_VAR
END_FUNCTION_BLOCK

METHOD ACT_02_PRODUCTIONSIMULATIONSETTINGS
END_METHOD

METHOD ACT_12_CALL_MACHINEPERFORMANCE
END_METHOD

METHOD ACT_00_BASE_CONVERSION
END_METHOD

METHOD ACT_01_STANDARDASSIGNMENTS
END_METHOD

METHOD ACT_11_BREAKASSIGNMENTS
END_METHOD

METHOD ACT_10_SCHEDULERSELECTION
END_METHOD

(* ---- L_OEEA_FBS.pou ---- *)
FUNCTION_BLOCK L_OEEA_FBS EXTENDS L_OEEA_FBs_COMMON
VAR_IN_OUT
	SCMACHINEDATA : scMachineData;
	SCPERFORMANCE : scPerformance;
	SCACTUALSTATEDURATION : scVisuProductionStatus_base;
	SCDOWNTIME : scDowntime;
	SCVISU_IN_X_TREND : scXAxis_Trend;
	SCVISU_IN_Y_TREND : scYAxis_Trend;
	SCVISU_TREND_Y_LIMITS : scTrend_Limits;
END_VAR
VAR
	FBMACHINEPERFORMANCE : L_OEEA_MachinePerformance;
	FBDOWNTIME : L_OEEA_Downtime;
	FB_X_AXIS_TREND : L_OEEA_X_TREND;
	FB_Y_AXIS_TREND : L_OEEA_Y_TREND;
	XSORTUPDOWN : BOOL := TRUE;
	FBTIMETRIGGER : TON;
	FBTIMETRIGGER2 : TON;
	TXYGRAPHTIME : TIME := TIME#1m0s0ms;
	SPOWERUPJSONSUBSTR : STRING(255);
	ISETCALCTHROUGHPUT : INT;
	TSETTIMEXYGRAPH : TIME;
END_VAR
END_FUNCTION_BLOCK

METHOD ACT_01_STANDARDASSIGNMENTS
END_METHOD

METHOD ACT_13_CALL_PRODUCTION_TRENDS
END_METHOD

METHOD ACT_02_PRODUCTIONSIMULATIONSETTINGS
END_METHOD

METHOD ACT_12_CALL_MACHINEPERFORMANCE
END_METHOD

METHOD ACT_11_BREAKASSIGNMENTS
END_METHOD

METHOD ACT_10_SCHEDULERSELECTION
END_METHOD

(* ---- L_OEEA_FBS_COMMON.pou ---- *)
FUNCTION_BLOCK L_OEEA_FBS_COMMON
VAR_INPUT
	XENABLED : BOOL;
	XRESETACTUALDATA : BOOL;
	XRESETHISTORYDATA : BOOL;
	XPRODSIMULTIONENABLED : BOOL;
	XPRODSIMEVENTOCCURRENCE : BOOL := TRUE;
	XPRODSIMMATERIALPRODUCTION : BOOL;
	XHMIACTIVE : BOOL;
	ESCHEDULERMODE : L_OEEA_BaseDependency.enumShiftMode;
	ESETWEEKDAY : RTCLK.WEEKDAY;
	XDEACTIVESHIFTCONTINIOUSUPDATE : BOOL;
	UIMAXSIMULATIONEVENTS : UINT := 1;
	SCTRIGGER : scTrigger;
	XUSERESONCODESTRING : BOOL;
	XUPDATEJSONOEEKPI : BOOL;
	XMANUALSHIFTRESET : BOOL;
	XSHIFTPRODUCTIONACTIVE : BOOL;
	XLATERSHIFTSTARTENABLED : BOOL;
	SCSIMULATIONMODES : scSimulationModes;
	SREASONTEXTPOWERON : STRING := '';
END_VAR
VAR_OUTPUT
	XBUSY : BOOL;
	XERROR : BOOL;
	SCSHIFTVALUES : L_OEEA_ShiftScheduler.scCurrentShiftValues;
END_VAR
VAR_IN_OUT
	SCPRODUCTIONMODE : scProductionMode;
	ASERRORCATEGORY : scCategoryStruct;
	SCFIRSTERRORDATA : scErrorData;
	ASCDAYSCHEDULES : ARRAY [1..uiDaySchedule] OF scDaySchedule;
	SCPDINTERNAL : scInternalVar;
	SCPDINTERNALDOWNTIME : scInternalDownVar;
	SCPDPRODUCTIONDATA : scInternalProductionData;
	SCPDSHIFTDAYINDEX : scPDShiftData;
	SCPDSHIFTHISTORY_BASE : scVisuShiftHistory_base;
	SCSHIFTDOWNTIMEHISTORY : ARRAY [1..3] OF scDowntime_base;
	SCOEE_VISUPD : scOEE_VisuPD;
	SCVISU_OUT_PARTCORRECTION : scPartCorrectionInput;
	SCVISU_OUT_BUTTONS : scVisuButtons;
	SCSIMULATIONDOWNTIMES : scSimulationDowntimes;
END_VAR
VAR
	FBOEEA_SIMULATIONSETTINGS : L_OEEA_SimulationSettings;
	FBPRODUCTIONSCHEDULER : L_OEEA_ProductionScheduler;
	SCCUTREAL : scCutAverageReal;
	FBSHIFTCALENDAR : L_OEEA_ShiftScheduler.L_OEEA_ShiftScheduler;
	FBSTANDARDASSIGNMENT : L_OEEA_StandardAssignment;
	FBSHIFTOEEHISTORY : L_OEEA_ShiftOEEHistory_base;
	EPRODLOGFORMAT : eProduction_log := eProduction_log.Json;
	FBSHIFTDOWNTIMEHISTORY : L_OEEA_ShiftDowntimeHistory_base;
	XFIRSTCYCLE : BOOL := FALSE;
	XGETDEACTIVESHIFTCONTINIOUSUPDATE : BOOL;
	SSHIFTNAME : STRING;
	ICALCTHROUGHPUT : INT := 0;
	XRESETPRODLOGSHIFTCHANGE : BOOL;
	XFIRSTPLCCYCLEPROLONG : BOOL;
	SETSHIFTNAME : scShiftName;
END_VAR
END_FUNCTION_BLOCK

(* ---- L_OEEA_LINE_FB.pou ---- *)
FUNCTION_BLOCK L_OEEA_LINE_FB
VAR_INPUT
	XENABLE : BOOL;
	XRESETHISTORY : BOOL;
	UIMAXNOOFMACHINES : UINT;
	UINOOFCONNCTEDMACHINES : UINT;
	UINOOFHISTORICALWEEKS : UINT;
	TSETTIMEDEVIATION : TIME := TIME#10s0ms;
	TSETTIMECONNECTION : TIME := TIME#1m30s0ms;
	TSETTIMESHIFTCHANGEDELAY : TIME := TIME#5s0ms;
	TSETTIMELINEOEEUPDATEDELAY : TIME := TIME#10s0ms;
	SCTRIGGER : scTrigger_base;
	SCMACHINEOFFMODE : scMachineOffMode;
	SSHIFTNAME : STRING;
	ILINEID : INT;
	SLINEID : STRING;
END_VAR
VAR_OUTPUT
	XBUSY : BOOL;
	XDONE : BOOL;
	XERROR : BOOL;
	SCLINESTATUS : scLineStatus;
	XSHIFTCHANGEDELAYPROLONGTIME : BOOL;
	XLINEOEEUPDATEDELAYPROLONGTIME : BOOL;
	XLINEOEESTORAGEDELAY : BOOL;
END_VAR
VAR_IN_OUT
	ASCMACHINEDATA_NVL : ARRAY [1..Line_OEE_GVL_Var.uiNoOfMachines] OF scMachineData_NVL;
	ASCNVL : ARRAY [1..Line_OEE_GVL_Var.uiNoOfMachines] OF scRef_NVL;
	SCSHIFTVALUES : scCurrentShiftValues;
	SCLINEKPIS : scLineKPIs;
	ASCHISTORICALLINEKPIS : ARRAY [1..Line_OEE_GVL_Var.uiNoOfHistoricalWeeks] OF scLineKPIs;
	SCACTIVEDURINGACTUALSHIFT : ARRAY [1..Line_OEE_GVL_Var.uiNoOfMachines] OF scMachineShiftActive;
END_VAR
VAR
	I : INT;
	K : INT;
	N : INT;
	SCLINEKPISDEL : scLineKPIs;
	SCLINESTATUSDEL : scLineStatus;
	ROEE_WEIGHT : REAL;
	ROEERT : REAL;
	RTEEP : REAL;
	SLASTDATETIME : STRING;
	DTLASTDATETIME : DATE_AND_TIME;
	ISTRPOSBLANK : INT;
	TDATETIMEDIFF : TIME;
	XFIRSTNOTCONNECTEDMACHINE : BOOL;
	XFIRSTMACHINEDATETIMEINSYNCH : BOOL;
	XFIRSTNOTACTIVEMACHINE : BOOL;
	DTSHIFTSTART : DATE_AND_TIME;
	IWEEKDAYSDIFF : INT;
	DTDIFFSTARTTIME : TIME;
	DTPREVIOUSDATETIME : DATE_AND_TIME;
	TONPROLONGTIMER : ARRAY [1..2] OF TON;
	ISTEPSHIFTCHANGE : INT := 0;
	XSHIFTCHANGELINECONTROLLERDETECTED : BOOL;
	ILASTNOMACHINEACTIVEOEECALC : INT;
	SCDELACTIVEDURINGACTUALSHIFT : ARRAY [1..Line_OEE_GVL_Var.uiNoOfMachines] OF scMachineShiftActive;
END_VAR
END_FUNCTION_BLOCK

METHOD ACT_LINEOEEHISTORY
END_METHOD

METHOD ACT_CAL_OEEKPIS
END_METHOD

METHOD ACT_SHIFTSTARTTIME
END_METHOD

METHOD SUB_01_INIT_LOOP
END_METHOD

METHOD SUB_02_CHECK_STATUS
END_METHOD

METHOD SUB_03_CALC_MACHINEOEE
END_METHOD

METHOD SUB_04_CALC_LINEOEESUMMARY
END_METHOD

METHOD SUB_05_CALC_AVERAGELINEOEE
END_METHOD

METHOD SUB_06_SET_LINESTATUS
END_METHOD

METHOD METH_PROLONGBIT : BOOL
VAR_INPUT
	TPROLONGTIME : TIME;
END_VAR
VAR_IN_OUT
	TONPROLONGTIMER : TON;
	XSTARTPROLONGTIME : BOOL;
END_VAR
END_METHOD

METHOD ACT_SHIFTCHANGESEQ
END_METHOD

(* ---- L_OEEA_SIMULATIONAXIS.pou ---- *)
FUNCTION_BLOCK L_OEEA_SIMULATIONAXIS
VAR_INPUT
	XENABLED : BOOL;
	XDOWNTIMESTOP : BOOL;
	RTECHNICALCYCLETIME : REAL;
END_VAR
VAR_OUTPUT
	XMANUALSTOP : BOOL;
END_VAR
VAR_IN_OUT
	LRAXESACTMETERS : LREAL;
	LRAXESACTSCAPMETERS : LREAL;
END_VAR
VAR
	AXISJOG : L_MC1A_BasicActuatingSpeed;
	XREGULATORON : BOOL;
	XMOVEVELEXECUTE : BOOL;
	XJOGPOS : BOOL;
	XSTOP : BOOL;
	LRJOGGINGSETVEL : LREAL;
	ISTEP : INT;
	RFACTORPERFORMANCELOSS : REAL := 1.025;
	LRACTUALINCPOSITIONSIM : LREAL;
	LRACTUALDIFF : LREAL;
	TSCRAPMATERIALSTART : TON_Pausable;
	TSCRAPMATERIALSTOP : TON_Pausable;
END_VAR
END_FUNCTION_BLOCK

METHOD ACTMOTIONCTRL
END_METHOD

METHOD ACT_CALLMOTIONFB
END_METHOD

(* ---- L_OEEA_SIMULATIONSETTINGS.pou ---- *)
FUNCTION_BLOCK L_OEEA_SIMULATIONSETTINGS
VAR_INPUT
	XPRODSIMULTIONENABLED : BOOL;
	XPRODSIMEVENTOCCURRENCE : BOOL := TRUE;
	XRESETACTUALDATA : BOOL;
	ESCHEDULERMODE : enumShiftMode;
	XMATERIALPRODUCTION : BOOL;
	UIMAXSIMULATIONEVENTS : UINT := 1;
	SCSIMULATIONMODES : scSimulationModes;
END_VAR
VAR_OUTPUT
	XBUSY : BOOL;
	XERROR : BOOL;
END_VAR
VAR_IN_OUT
	SCMACHINEDATA : scMachineData;
	SCSHIFTVALUES : L_OEEA_ShiftScheduler.scCurrentShiftValues;
	SCDOWNTIME : scDowntime;
	SCSIMULATIONDOWNTIMES : scSimulationDowntimes;
	SCPRODUCTIONMODE : scProductionMode;
END_VAR
VAR
	SCRT_STATUS : RT_Status_Struct;
	FBDATASIMULATOR : L_OEEA_DataSimulator;
	XSTATIONENABLED : BOOL := TRUE;
	SCRT_STATUS_RESET : RT_Status_Struct;
	PA_TIMER : RT_Timer;
	PA_DOWNTIME : RT_Downtime;
	SCCUTREAL : scCutAverageReal;
	XFIRSTCYCLESIM : BOOL := FALSE;
	FBXHOLDINGACTIVE : R_TRIG;
	DILASTTYPEID : INT;
	IMAXSIMULATIONERRORS : INT;
	FBSIMULATIONAXIS : L_OEEA_SimulationAxis;
	XMANUALSTOP : BOOL;
	LRCOUNTOK : LREAL;
	LRCOUNTNOK : LREAL;
END_VAR
END_FUNCTION_BLOCK

METHOD ACT_03_MASCHINEPERFORMANCESIMULATION
END_METHOD

METHOD ACT_01_PRODUCTIONSIMULATION
END_METHOD

METHOD ACT_02_CALL_PRODUCTIONSIMULATOR
END_METHOD

METHOD ACT_04_CALLSIMULATIONAXIS
END_METHOD

(* ---- L_OEEA_STANDARDASSIGNMENT.pou ---- *)
FUNCTION_BLOCK L_OEEA_STANDARDASSIGNMENT
VAR_INPUT
	ENABLED : BOOL;
	XHMIACTIVE : BOOL;
END_VAR
VAR_OUTPUT
	XBUSY : BOOL;
	XERROR : BOOL;
END_VAR
VAR_IN_OUT
	SCSHIFTVALUES : L_OEEA_ShiftScheduler.scCurrentShiftValues;
	SCMACHINEDATA : scMachineData;
	SCDOWNTIME : scDowntime;
	SCPRODUCTIONMODE : scProductionMode;
	ASERRORCATEGORY : scCategoryStruct;
	SCFIRSTERRORDATA : scErrorData;
	ASCDAYSCHEDULES : ARRAY [1..uiDaySchedule] OF scDaySchedule;
	SCOEE_VISUPD : scOEE_VisuPD;
	SCVISU_OUT_BUTTONS : scVisuButtons;
	SCVISU_OUT_PARTCORRECTION : scPartCorrectionInput;
END_VAR
VAR
	I : INT;
	K : INT;
	IDEFAULTDAYOFWEEK : INT;
	IACTUALDAYOFWEEK : INT;
	XFIRSTCYCLE : BOOL := FALSE;
	FBXSAVESHIFTDATA : R_TRIG;
	ACTUALDAYINDEX : INT;
END_VAR
END_FUNCTION_BLOCK

METHOD ACT_01_PRODUCTIONMODES
END_METHOD

METHOD ACT_02_SETSHIFTINTERVALS
END_METHOD

METHOD ACT_03_MACHINEPERFORMANCESETTINGS
END_METHOD

(* ---- L_OEEA_VALIDATION_FBS.pou ---- *)
FUNCTION_BLOCK L_OEEA_VALIDATION_FBS EXTENDS L_OEEA_FBs
VAR
	FBPRODUCTIONSCHEDULER2 : L_OEEA_ProductionScheduler;
END_VAR
END_FUNCTION_BLOCK

METHOD ACT_12X_CALL_MACHINEPERFROMANCETEST
END_METHOD

(* ---- L_TB1A_PT1FILTER.pou ---- *)
FUNCTION_BLOCK L_TB1A_PT1FILTER
VAR_INPUT
	LRIN : LREAL;
	LRFILTERTIME : LREAL := 0.1;
END_VAR
VAR_OUTPUT
	LROUT : LREAL;
END_VAR
VAR
	TON0 : TON := STRUCT(IN := TRUE, PT := TIME#1m0s0ms);
	X1STCYCLE : BOOL := TRUE;
	BYINITCOUNTER : BYTE;
	LRTASKCYCLETIME : LREAL;
END_VAR
END_FUNCTION_BLOCK
